(* IEC 61131-3 sources: guidance-for-physical-ai-production-designer-on-aws/source/plan2cell/examples/welding_cell_2_small/plc/codesys/head/POU, 8 files *)

(* ---- FB_Cell.st ---- *)
(*
 * FB_Cell
 * Generated by bt2plc 0.1.0 for cell welding_cell_2_small (plan bt_1790934549_welding_cell_2_small)
 *
 * Cell control for 2 robot(s): bring-up, blind homing (HOME_FOLGE), production
 * cycle (awRobotProdFolge started on every active robot; the robots run autonomously),
 * zone / permit arbitration (FB_ZoneArbiter), supervision (op index sequence, per-op
 * watchdog, zone-wait deadline, stall, program completeness), abort (stop all, drop grants,
 * rewind tickets), recovery confirmation and reset (Reset held >= 500 ms).
 *
 *   INIT -> BRINGUP -> HOMING_SELECT <-> HOMING_RUN -> READY -> START_JOBS -> RUNNING
 *        -> CYCLE_DONE -> READY ...
 *   any fault -> ABORTING -> ERROR -(bReset)-> RESETTING -> BRINGUP -> HOMING_SELECT ...
 *   abort with a robot inside its program (op index > 0, grant held, program left
 *   incomplete or away from home), or the first bring-up after INIT (head restart /
 *   download) with an active robot away from home:
 *        ... BRINGUP -> RECOVERY -(bRecoveryConfirm)-> RESETTING -> BRINGUP -> HOMING_SELECT
 *        (operator moves the robots clear in T1 first; homing is then always sequential)
 *   Start-up homing stays automatic when every active robot is at home.
 *
 * Operator: a bStop edge is latched in every state until it is consumed - abort (normal
 * states), cancel of the reset -> ERROR (INIT / RESETTING, driver Reset low), or cleared
 * (ERROR). A bReset edge in ABORTING is applied when ERROR is reached.
 *
 * Scan order: robot drivers (commands of the previous scan) -> op index tracking ->
 * faults known so far -> arbiter (this scan's inputs, no new grants after a fault) ->
 * watchdogs -> faults -> state machine -> GRANT bytes (0 when a fault is latched).
 * Op supervision runs whenever a robot's production job is commanded / running, in any
 * cell state: op index sequence, zone ops left without grant, op index 0 while running.
 *
 * Portable: one FB_VassRobot instance per robot (no FB instance arrays), timers are
 * TIME stamps of one free-running clock (_tNow).
 *)

FUNCTION_BLOCK FB_Cell
VAR_INPUT
    bEnable             : BOOL := TRUE;
    bAutoRun            : BOOL := TRUE;     (* Level: start a cycle whenever READY *)
    bStart              : BOOL;             (* Rising edge: start one cycle *)
    bStop               : BOOL;             (* Rising edge: abort (ERR_OPERATOR_STOP) *)
    bReset              : BOOL;             (* Rising edge in CS_ERROR: reset robots and cell *)
    bRecoveryConfirm    : BOOL;             (* Rising edge (from CS_ERROR on, while bRecoveryRequired): robots cleared *)
    astIn               : ARRAY[1..2] OF ST_RobotIn;    (* Robot inputs (copied from GVL_IO) *)
END_VAR

VAR_OUTPUT
    astOut              : ARRAY[1..2] OF ST_RobotOut;   (* Robot outputs (copied to GVL_IO) *)
    eState              : E_CellState;
    eError              : E_CellError;      (* First fault, ERR_NONE when OK *)
    nErrorRobot         : INT;              (* Robot of the fault, 0 = cell *)
    nErrorOp            : INT;              (* Op index of the fault, 0 = none *)
    nErrorZone          : INT;              (* Zone of the fault, 0 = none *)
    bCycleActive        : BOOL;             (* START_JOBS or RUNNING *)
    bError              : BOOL;             (* Fault latched until the reset is done *)
    bHomingRequired     : BOOL;         (* Profile vw-ks24: a robot is not at home and must be
                                           jogged there by the operator (no blind HOME Folge) *)
    bRecoveryRequired   : BOOL;             (* bRecoveryConfirm needed before homing (abort mid-cycle / start-up away from home) *)
    udiCycles           : UDINT;            (* Completed production cycles *)
    tLastCycle          : TIME;             (* Duration of the last cycle (RUNNING) *)
    aeRobotState        : ARRAY[1..2] OF E_RobotState;
    aeRobotError        : ARRAY[1..2] OF E_CellError;
    awStep              : ARRAY[1..2] OF WORD;          (* Reported op index *)
    adwReq              : ARRAY[1..2] OF DWORD;         (* REQUEST per robot *)
    adwGrant            : ARRAY[1..2] OF DWORD;         (* GRANT per robot (as sent) *)
    anDone              : ARRAY[1..2] OF INT;           (* Ops completed in this cycle *)
    anHolder            : ARRAY[1..2] OF INT;        (* Zone holder, 0 = free *)
    anTicket            : ARRAY[1..2] OF INT;        (* Next ticket per zone *)
END_VAR

VAR
    (* ========================================================================
       ROBOT DRIVERS (one instance per robot) AND ARBITER
       ======================================================================== *)
    fbRobot_R1          : FB_VassRobot;     (* 1: robot1 - kuka_robi1 (192.168.100.11) *)
    fbRobot_R2          : FB_VassRobot;     (* 2: robot2 - kuka_robi2 (192.168.100.12) *)
    fbArbiter           : FB_ZoneArbiter;

    (* ========================================================================
       CELL STATE
       ======================================================================== *)
    _eState             : E_CellState := E_CellState.CS_INIT;
    _eLastState         : E_CellState := E_CellState.CS_INIT;
    _bFault             : BOOL;             (* Fault latched (eError valid) *)
    _bPowerOn           : BOOL;             (* Robots: bring up *)
    _bArbReset          : BOOL := TRUE;     (* Arbiter reset in the next scan *)
    _bNeedRecovery      : BOOL;             (* Latched at an abort with a robot inside its program *)
    _bRecoveryHoming    : BOOL;             (* Homing after recovery: always sequential *)
    _bEngaged           : BOOL;             (* A robot is inside its production program / holds a grant *)
    _bConfirmLatch      : BOOL;             (* bRecoveryConfirm edge seen since CS_ERROR *)
    _bFirstBringup      : BOOL := TRUE;     (* First bring-up after CS_INIT: check the home poses *)
    _bStopReq           : BOOL;             (* bStop edge, latched until consumed *)
    _bResetReq          : BOOL;             (* bReset edge seen in CS_ABORTING, applied in CS_ERROR *)
    _bFaultScan         : BOOL;             (* Fault source known before the arbiter call (this scan) *)

    (* ========================================================================
       ROBOT STATUS (copied from the driver instances every scan)
       ======================================================================== *)
    _abIdle             : ARRAY[1..2] OF BOOL;
    _abBusy             : ARRAY[1..2] OF BOOL;
    _abDrvError         : ARRAY[1..2] OF BOOL;          (* Driver in RS_ERROR / RS_RESET *)
    _abJobActive        : ARRAY[1..2] OF BOOL;
    _abJobDone          : ARRAY[1..2] OF BOOL;
    _abAtHome           : ARRAY[1..2] OF BOOL;
    _abRobotError       : ARRAY[1..2] OF BOOL;          (* Robot reports Error *)
    _abProgRunning      : ARRAY[1..2] OF BOOL;          (* Robot reports ProgRunning *)
    _awLastStep         : ARRAY[1..2] OF WORD;

    (* ========================================================================
       COMMANDS TO THE ROBOT DRIVERS (used in the next scan)
       ======================================================================== *)
    _abJobCmd           : ARRAY[1..2] OF BOOL;
    _awJob              : ARRAY[1..2] OF WORD;
    _abProdCmd          : ARRAY[1..2] OF BOOL;          (* Commanded job is the production Folge *)
    _abStopCmd          : ARRAY[1..2] OF BOOL;
    _abResetCmd         : ARRAY[1..2] OF BOOL;
    _abHoming           : ARRAY[1..2] OF BOOL;

    (* ========================================================================
       PRODUCTION CYCLE SUPERVISION
       ======================================================================== *)
    _abHasJob           : ARRAY[1..2] OF BOOL;          (* Active robot with ops *)
    _abRobotOk          : ARRAY[1..2] OF BOOL;          (* Arbiter input *)
    _anDone             : ARRAY[1..2] OF INT;           (* Arbiter input: ops completed *)
    _anStepSeen         : ARRAY[1..2] OF INT;           (* Op index seen last scan (incl. 0) *)
    _anLastStep         : ARRAY[1..2] OF INT;           (* Last validated non-zero op index *)
    _abGranted          : ARRAY[1..2] OF BOOL;          (* Current zone op has been granted *)
    _abOpRun            : ARRAY[1..2] OF BOOL;          (* Op watchdog running *)
    _atOpStart          : ARRAY[1..2] OF TIME;
    _abStallRun         : ARRAY[1..2] OF BOOL;          (* Stall watchdog running *)
    _atStallStart       : ARRAY[1..2] OF TIME;
    _abZeroRun          : ARRAY[1..2] OF BOOL;          (* Op index 0 watchdog running *)
    _atZeroStart        : ARRAY[1..2] OF TIME;
    _tCycleStart        : TIME;

    (* ========================================================================
       TIME BASE / TIMERS / EDGES
       ======================================================================== *)
    _tonClock           : TON;              (* Free-running clock, restarted every hour *)
    _tClockBase         : TIME;
    _tNow               : TIME;             (* Monotonic time of this scan *)
    _tonState           : TON;              (* State timeout, restarts on every state change *)
    _tLimit             : TIME;
    _rtrigStart         : R_TRIG;
    _rtrigStop          : R_TRIG;
    _rtrigReset         : R_TRIG;
    _rtrigConfirm       : R_TRIG;

    (* ========================================================================
       SCRATCH
       ======================================================================== *)
    _eNew               : E_CellError;
    _nNewRobot          : INT;
    _nNewOp             : INT;
    _nHomeCount         : INT;
    _nDone              : INT;
    _r                  : INT;
    _iOp                : INT;
    _nStep              : INT;
    _nPrev              : INT;              (* Op index that is left *)
    _tZeroLimit         : TIME;
    _dwGrant            : DWORD;
    _bBypass            : BOOL;
    _bAll               : BOOL;
    _bSequential        : BOOL;

    (* Profile vw-ks24: interlock grant / partner release encoding *)
    _z                  : INT;
    _q                  : INT;
    _nIl                : INT;
    _nIlQ               : INT;
    _nIdx               : INT;
    _nB                 : INT;
    _nBit               : INT;
    _wBits              : WORD;
    _bGrantBit          : BOOL;
    _bPartner           : BOOL;
END_VAR

(* ---- FB_VassRobot.st ---- *)
(*
 * FB_VassRobot
 * Generated by bt2plc 0.1.0 for cell welding_cell_2_small (plan bt_1790934549_welding_cell_2_small)
 *
 * VW VASS protocol driver for ONE robot (KUKA VKRC nexxt V8.2 DIM 2 via PROFINET).
 * Portable: no pointers, no REFERENCE, no OOP - the robot IO is passed as struct
 * copies (stIn / stOut) by the caller (FB_Cell, PLC_PRG copies GVL_IO).
 *
 *   Bring-up : SAFETY_ENABLE (T_BRINGUP_LIMIT: PROFINET / PROFIsafe connection set-up)
 *              -> DRIVES_ON -> MODE_EXT -> IDLE   (T_HANDSHAKE each)
 *   Job      : WAIT_READY -> SEND (echo checked) -> START (T_START_PULSE) -> WAIT_RUNNING
 *              -> RUNNING -> DONE   (WAIT_RUNNING -> DONE if the job finished between scans)
 *              (RUNNING -> ERROR ERR_ROBOT_STOPPED only after ProgRunning and ProgFinished
 *              stayed low for T_STOP_DEBOUNCE: a robot may publish the two bits in different
 *              bus frames at the Folge end)
 *              (T_HANDSHAKE per handshake state)
 *   Abort    : STOPPING (Stop + Cancel held >= T_STOP_PULSE and until ProgRunning drops)
 *   Recovery : ERROR -> RESET (Reset held T_RESET_PULSE >= 500 ms while bCmdReset stays TRUE;
 *              bCmdReset dropped = reset cancelled -> ERROR) -> SAFETY_ENABLE
 *              (still ProgRunning after the pulse -> ERROR, ERR_STOP_TIMEOUT)
 *   Command handshake: bCmdJob is a level request (rising edge latched),
 *              bJobDone the acknowledge (cleared while bCmdJob = FALSE).
 *
 * Stop is never dropped while the robot still reports ProgRunning (also in ERROR / RESET).
 * ProgRunning outside a job (OFF, bring-up, IDLE) -> ERROR (ERR_UNEXPECTED_RUN, Stop + Cancel).
 * The zone GRANT bytes (GVL_Cell.GRANT_BYTE .. +3) are written 0 here: FB_Cell encodes
 * them after FB_ZoneArbiter has run, so a grant reaches the robot in the scan it is computed.
 *
 * Profile vw-ks24 (GVL_Cell.PROFILE_VW): the VW tech package on the robot does the Folge
 * handshake, so the signal map and the job states differ (same state names):
 *   status  : ready A9, safety A10 + A13, auto A12, home A15 (PF0), Folge end A14,
 *             echo PRG_NR_REFL A1-8, op index P_PktNr_SPS, error code VW_FEH_BIN_A
 *   commands: drives E10, Folge number PRG_NR E1-8, start SRB E9 (level), reset E26
 *   job     : SEND writes PRG_NR and waits for the echo; START holds SRB until the robot
 *             leaves home (its cycle-start point clears PF0); RUNNING waits for Folge end;
 *             DONE clears PRG_NR and waits for the Folge end to fall
 *   zones   : REQUEST bit z is synthesised as "requesting or occupying",
 *             A(80+n) OR NOT A(40+n), which is exactly the REQUEST semantics of the arbiter;
 *             the release is A(40+n) going TRUE again. There is no 4-phase handshake.
 *   stop    : no Stop/Cancel bits exist; the head drops the drives, withdraws the partner
 *             releases (the robot's online driving condition stops it on the path) and clears
 *             PRG_NR. Recovery needs manual homing (PF0), there is no blind HOME Folge.
 *)

FUNCTION_BLOCK FB_VassRobot
VAR_INPUT
    bEnable             : BOOL := TRUE;
    nRobot              : INT := 1;         (* 1-based robot index (profile vw-ks24: interlock map) *)
    bPowerOn            : BOOL;             (* Level: bring the robot up *)
    bCmdJob             : BOOL;             (* Level request (rising edge latched): run job wJobNr *)
    wJobNr              : WORD;             (* Folge number, latched at job accept *)
    bProdJob            : BOOL;             (* wJobNr is the production Folge: send PLAN_ID, track wLastStep *)
    bCmdStop            : BOOL;             (* Level: abort the active job *)
    bCmdReset           : BOOL;             (* Rising edge in RS_ERROR: reset the robot; hold until bError drops *)
    stIn                : ST_RobotIn;       (* Copy of this robot's GVL_IO inputs *)
END_VAR

VAR_OUTPUT
    stOut               : ST_RobotOut;      (* Copy to this robot's GVL_IO outputs (GRANT bytes = 0) *)
    eState              : E_RobotState;
    eError              : E_CellError;
    bIdle               : BOOL;
    bBusy               : BOOL;             (* Job, stopping or resetting *)
    bJobActive          : BOOL;             (* Job started and ProgRunning *)
    bJobDone            : BOOL;             (* Job finished (cleared while bCmdJob = FALSE) *)
    bError              : BOOL;             (* RS_ERROR or RS_RESET *)

    (* Decoded robot status *)
    bDrivesOn           : BOOL;
    bProgRunning        : BOOL;
    bAtHome             : BOOL;
    bModeExt            : BOOL;
    bRobotReady         : BOOL;
    bRobotError         : BOOL;
    bProgFinished       : BOOL;
    bJobAck             : BOOL;
    bSafetyOK           : BOOL;
    wActiveJob          : WORD;             (* Echoed job number *)
    wStep               : WORD;             (* Reported op index, 0 = no program *)
    wLastStep           : WORD;             (* Max op index of the running production job (cleared at job accept) *)
    dwZoneReq           : DWORD;            (* REQUEST DWORD: zone bits 0..30, permit bit 31 *)
    wRobotErrorCode     : WORD;
END_VAR

VAR
    _eState             : E_RobotState := E_RobotState.RS_OFF;
    _eLastState         : E_RobotState := E_RobotState.RS_OFF;
    _wJob               : WORD;             (* Job number latched at accept *)
    _bProdJob           : BOOL;             (* Latched bProdJob *)
    _bJobPending        : BOOL;             (* Job edge seen, not yet accepted *)
    _bInJob             : BOOL;
    _bUp                : BOOL;
    _bNoJob             : BOOL;             (* Off / bring-up / idle: ProgRunning is not expected *)

    (* Commands to the robot *)
    _bSafeEnable        : BOOL;
    _bDrivesOnCmd       : BOOL;
    _bExtCmd            : BOOL;
    _bStartCmd          : BOOL;
    _bStopCmd           : BOOL;
    _bCancelCmd         : BOOL;
    _bResetCmd          : BOOL;
    _bJobReqCmd         : BOOL;

    (* Timers *)
    _tonStep            : TON;              (* State timeout, restarts on every state change *)
    _tonPulse           : TON;              (* Start / stop / reset pulse width *)
    _tonStopDebounce    : TON;              (* RS_JOB_RUNNING: ProgRunning + ProgFinished low (T_STOP_DEBOUNCE) *)
    _tStepLimit         : TIME;

    (* Edge detection *)
    _rtrigJob           : R_TRIG;
    _rtrigReset         : R_TRIG;

    (* Profile vw-ks24 *)
    _bFolgeEnd          : BOOL;             (* A14 Folge end *)
    _bVwStarted         : BOOL;             (* SRB acknowledged: the robot left its home point *)
    _nIdx               : INT;              (* signal index 1..256 *)
    _nB                 : INT;              (* telegram byte of _nIdx *)
    _nBit               : INT;              (* bit of _nIdx *)
    _wTmp               : WORD;
    _bTmp               : BOOL;
    _z                  : INT;
    _n                  : INT;

    _i                  : INT;
END_VAR

(* ---- FB_ZoneArbiter.st ---- *)
(*
 * FB_ZoneArbiter
 * Generated by bt2plc 0.1.0 for cell welding_cell_2_small (plan bt_1790934549_welding_cell_2_small)
 *
 * Zone (mutex) and permit arbiter, data-driven by GVL_Cell (aTickets, anZoneFirst/Count,
 * aOps[].dwZoneMask / nPredFirst / nPredCount, aPreds).
 *
 * REQUEST / GRANT DWORD: bits 0..30 = zones 1..31, bit 31 = PERMIT (GVL_Cell.PERMIT_MASK).
 *   GP_PLANNED : a zone is granted only to its next ticket holder, only if the request
 *                equals the op's full mask and the reported op index matches the ticket.
 *   GP_FCFS    : free zones to any requester whose request equals the op mask, oldest
 *                request first, ties by robot index; zones of an older requester that
 *                waits only for occupied zones are reserved against younger ones.
 *                BT ordering is NOT preserved by the zones.
 *   PERMIT     : granted for op (r, k) iff every pred (q, j) of the op has anDone[q] >= j.
 *                Not a mutex: never held against other robots, released when bit 31 drops.
 * Both policies grant all bits of an op in the same scan (all-or-nothing).
 *
 * Checks: 4-phase handshake (op index must not change while a grant is held), release
 * only by a robot that runs OK, holder raising extra bits; request mask and ticket checks
 * are evaluated once (op index, REQUEST) has been stable for tDebounce.
 * Fail closed: any violation latches bFault and drops all grants until bReset.
 *
 * Timing uses tNow (monotonic TIME from the caller's clock), no timer instances.
 *)

FUNCTION_BLOCK FB_ZoneArbiter
VAR_INPUT
    bReset              : BOOL;             (* Level: rewind tickets, clear holders, grants and fault *)
    bEnable             : BOOL;             (* New grants allowed *)
    ePolicy             : E_GrantPolicy := E_GrantPolicy.GP_PLANNED;
    tDebounce           : TIME := T#200MS;  (* (op index, REQUEST) stable time before mask / ticket checks *)
    tNow                : TIME;             (* Monotonic time of this scan *)
    abRobotOk           : ARRAY[1..2] OF BOOL;      (* Production job running, no robot error *)
    awStep              : ARRAY[1..2] OF WORD;      (* Reported op index, 0 = none *)
    adwReq              : ARRAY[1..2] OF DWORD;     (* REQUEST DWORD *)
    anDone              : ARRAY[1..2] OF INT;       (* Ops completed per robot in this cycle *)
END_VAR

VAR_OUTPUT
    adwGrant            : ARRAY[1..2] OF DWORD;     (* GRANT DWORD per robot *)
    anHolder            : ARRAY[1..2] OF INT;    (* Robot holding the zone, 0 = free *)
    anTicket            : ARRAY[1..2] OF INT;    (* Next ticket index in GVL_Cell.aTickets *)
    bAllConsumed        : BOOL;             (* No zone held and (planned) every ticket consumed *)
    bFault              : BOOL;
    eFault              : E_CellError;
    nFaultRobot         : INT;
    nFaultZone          : INT;
END_VAR

VAR
    _udiScan            : UDINT;            (* Scan counter: request age for FCFS *)
    _audiWaitSince      : ARRAY[1..2] OF UDINT;     (* Scan of the first pending request, 0 = none *)
    _abPicked           : ARRAY[1..2] OF BOOL;
    _anGrantStep        : ARRAY[1..2] OF INT;       (* Op index at the time of the grant *)
    _awPrevStep         : ARRAY[1..2] OF WORD;
    _adwPrevReq         : ARRAY[1..2] OF DWORD;
    _atChange           : ARRAY[1..2] OF TIME;      (* tNow of the last (op index, REQUEST) change *)
    _abStable           : ARRAY[1..2] OF BOOL;
    _eNew               : E_CellError;
    _nNewRobot          : INT;
    _nNewZone           : INT;
    _k                  : INT;
    _r                  : INT;
    _rr                 : INT;
    _rSel               : INT;
    _z                  : INT;
    _p                  : INT;
    _q                  : INT;
    _iOp                : INT;
    _nStep              : INT;
    _nTicket            : INT;
    _nLastTicket        : INT;
    _nPredFirst         : INT;
    _nPredLast          : INT;
    _dwBit              : DWORD;
    _dwExp              : DWORD;            (* Expected REQUEST of the reported op *)
    _dwZones            : DWORD;            (* Zone bits of _dwExp (permit bit removed) *)
    _dwReserved         : DWORD;            (* FCFS: zones reserved by older requesters this scan *)
    _bOk                : BOOL;             (* All zones of the op grantable *)
    _bPermitOk          : BOOL;             (* All permit predecessors done *)
    _bPending           : BOOL;
END_VAR

(* ---- FB_Cell_Body.st ---- *)
(*
 * FB_Cell - Implementation
 *)

IF NOT bEnable THEN
    _eState := E_CellState.CS_INIT;
END_IF

(* ============================================================================
   TIME BASE / EDGES
   ============================================================================ *)
_tonClock(IN := TRUE, PT := T#1H);
_tNow := _tClockBase + _tonClock.ET;
IF _tonClock.Q THEN
    _tClockBase := _tNow;
    _tonClock(IN := FALSE);
    _tonClock(IN := TRUE, PT := T#1H);
END_IF

_rtrigStart(CLK := bStart);
_rtrigStop(CLK := bStop);
_rtrigReset(CLK := bReset);
_rtrigConfirm(CLK := bRecoveryConfirm);

(* Operator stop: latched in every state until consumed (abort, cancelled reset, CS_ERROR);
   it also cancels a reset that is pending from CS_ABORTING *)
IF _rtrigStop.Q THEN
    _bStopReq := TRUE;
    _bResetReq := FALSE;
END_IF

FOR _r := 1 TO GVL_Cell.N_ROBOTS DO
    _abHasJob[_r] := GVL_Cell.abRobotActive[_r] AND (GVL_Cell.anRobotOpCount[_r] > 0);
END_FOR

(* ============================================================================
   ROBOT DRIVERS (commands from the previous scan; GRANT bytes are added below)
   ============================================================================ *)

(* 1: R1 - robot1 *)
fbRobot_R1(
    bEnable     := bEnable,
    bPowerOn    := _bPowerOn,
    bCmdJob     := _abJobCmd[1],
    wJobNr      := _awJob[1],
    bProdJob    := _abProdCmd[1],
    bCmdStop    := _abStopCmd[1],
    bCmdReset   := _abResetCmd[1],
    nRobot      := 1,
    stIn        := astIn[1]);
astOut[1]         := fbRobot_R1.stOut;
aeRobotState[1]   := fbRobot_R1.eState;
aeRobotError[1]   := fbRobot_R1.eError;
awStep[1]         := fbRobot_R1.wStep;
adwReq[1]         := fbRobot_R1.dwZoneReq;
_awLastStep[1]    := fbRobot_R1.wLastStep;
_abIdle[1]        := fbRobot_R1.bIdle;
_abBusy[1]        := fbRobot_R1.bBusy;
_abDrvError[1]    := fbRobot_R1.bError;
_abJobActive[1]   := fbRobot_R1.bJobActive;
_abJobDone[1]     := fbRobot_R1.bJobDone;
_abAtHome[1]      := fbRobot_R1.bAtHome;
_abRobotError[1]  := fbRobot_R1.bRobotError;
_abProgRunning[1] := fbRobot_R1.bProgRunning;

(* 2: R2 - robot2 *)
fbRobot_R2(
    bEnable     := bEnable,
    bPowerOn    := _bPowerOn,
    bCmdJob     := _abJobCmd[2],
    wJobNr      := _awJob[2],
    bProdJob    := _abProdCmd[2],
    bCmdStop    := _abStopCmd[2],
    bCmdReset   := _abResetCmd[2],
    nRobot      := 2,
    stIn        := astIn[2]);
astOut[2]         := fbRobot_R2.stOut;
aeRobotState[2]   := fbRobot_R2.eState;
aeRobotError[2]   := fbRobot_R2.eError;
awStep[2]         := fbRobot_R2.wStep;
adwReq[2]         := fbRobot_R2.dwZoneReq;
_awLastStep[2]    := fbRobot_R2.wLastStep;
_abIdle[2]        := fbRobot_R2.bIdle;
_abBusy[2]        := fbRobot_R2.bBusy;
_abDrvError[2]    := fbRobot_R2.bError;
_abJobActive[2]   := fbRobot_R2.bJobActive;
_abJobDone[2]     := fbRobot_R2.bJobDone;
_abAtHome[2]      := fbRobot_R2.bAtHome;
_abRobotError[2]  := fbRobot_R2.bRobotError;
_abProgRunning[2] := fbRobot_R2.bProgRunning;

(* A robot inside its production program or holding a grant (previous scan's commands):
   inside an op, between two ops, finished with an incomplete program, or left the
   home pose during the current cycle *)
_bEngaged := FALSE;
FOR _r := 1 TO GVL_Cell.N_ROBOTS DO
    IF _abJobCmd[_r] AND _abProdCmd[_r] THEN
        IF awStep[_r] <> WORD#0 THEN
            _bEngaged := TRUE;
        ELSIF (_awLastStep[_r] <> WORD#0) AND NOT _abJobDone[_r] THEN
            _bEngaged := TRUE;
        ELSIF _abJobDone[_r] AND (WORD_TO_INT(_awLastStep[_r]) <> GVL_Cell.anRobotOpCount[_r]) THEN
            _bEngaged := TRUE;
        ELSIF NOT _abAtHome[_r]
              AND ((_awLastStep[_r] <> WORD#0) OR (_anLastStep[_r] <> 0) OR _abJobActive[_r]) THEN
            _bEngaged := TRUE;
        END_IF
    END_IF
    IF fbArbiter.adwGrant[_r] <> DWORD#0 THEN
        _bEngaged := TRUE;
    END_IF
END_FOR

(* ============================================================================
   OP INDEX TRACKING (production job commanded, any cell state)
   The index must advance by exactly +1. The op that is left (also at the job end,
   index -> 0) must have been granted if it has a zone / permit mask (both policies).
   Index 0 while the program runs is valid only before the first / after the last op.
   ============================================================================ *)
_eNew := E_CellError.ERR_NONE;
_nNewRobot := 0;
_nNewOp := 0;
FOR _r := 1 TO GVL_Cell.N_ROBOTS DO
    IF _abJobCmd[_r] AND _abProdCmd[_r] THEN
        _nStep := WORD_TO_INT(awStep[_r]);
        IF _nStep <> _anStepSeen[_r] THEN
            _nPrev := _anStepSeen[_r];
            _bBypass := FALSE;
            IF (_nPrev >= 1) AND (_nPrev <= GVL_Cell.anRobotOpCount[_r]) AND NOT _abGranted[_r] THEN
                _iOp := GVL_Cell.anRobotFirstOp[_r] + _nPrev - 1;
                IF GVL_Cell.aOps[_iOp].dwZoneMask <> DWORD#0 THEN
                    _bBypass := TRUE;               (* zone / permit op left without a grant *)
                END_IF
            END_IF
            IF _bBypass THEN
                IF _eNew = E_CellError.ERR_NONE THEN
                    _eNew := E_CellError.ERR_ZONE_BYPASSED;
                    _nNewRobot := _r;
                    _nNewOp := _nPrev;
                END_IF
            ELSIF _nStep <> 0 THEN
                IF (_nStep = _anLastStep[_r] + 1) AND (_nStep <= GVL_Cell.anRobotOpCount[_r]) THEN
                    _anLastStep[_r] := _nStep;
                ELSIF _eNew = E_CellError.ERR_NONE THEN
                    _eNew := E_CellError.ERR_STEP_SEQUENCE;
                    _nNewRobot := _r;
                    _nNewOp := _nStep;
                END_IF
            END_IF
            _anStepSeen[_r] := _nStep;
            _abGranted[_r] := FALSE;
            _abOpRun[_r] := FALSE;
            _abStallRun[_r] := FALSE;
            _abZeroRun[_r] := FALSE;
        END_IF

        (* index 0 while the program runs, between two ops *)
        IF _abJobActive[_r] AND (_nStep = 0) AND (_anLastStep[_r] > 0)
           AND (_anLastStep[_r] < GVL_Cell.anRobotOpCount[_r])
           AND (_eNew = E_CellError.ERR_NONE) THEN
            _eNew := E_CellError.ERR_STEP_SEQUENCE;
            _nNewRobot := _r;
            _nNewOp := 0;
        END_IF

        (* ops completed (permit predecessors): validated index - 1, all at job done *)
        IF _abJobDone[_r] AND (_anLastStep[_r] = GVL_Cell.anRobotOpCount[_r]) THEN
            _nDone := GVL_Cell.anRobotOpCount[_r];
        ELSIF _anLastStep[_r] > 0 THEN
            _nDone := _anLastStep[_r] - 1;
        ELSE
            _nDone := 0;
        END_IF
        _anDone[_r] := MAX(_anDone[_r], _nDone);
    END_IF
END_FOR

(* ============================================================================
   ZONE ARBITER (this scan's robot inputs)
   No new grants in a scan in which the cell already knows it will abort:
   driver error, latched operator stop, latched fault, supervision fault above.
   ============================================================================ *)
_bFaultScan := _bFault OR _bStopReq OR (_eNew <> E_CellError.ERR_NONE);
FOR _r := 1 TO GVL_Cell.N_ROBOTS DO
    _abRobotOk[_r] := _abJobActive[_r] AND _abJobCmd[_r] AND _abProdCmd[_r] AND NOT _abRobotError[_r];
    IF _abDrvError[_r] THEN
        _bFaultScan := TRUE;
    END_IF
END_FOR
fbArbiter(
    bReset      := _bArbReset,
    bEnable     := ((_eState = E_CellState.CS_START_JOBS) OR (_eState = E_CellState.CS_RUNNING))
                   AND NOT _bFaultScan,
    ePolicy     := GVL_Cell.GRANT_POLICY,
    tDebounce   := GVL_Cell.T_MISMATCH_DEBOUNCE,
    tNow        := _tNow,
    abRobotOk   := _abRobotOk,
    awStep      := awStep,
    adwReq      := adwReq,
    anDone      := _anDone);
_bArbReset := FALSE;

(* ============================================================================
   WATCHDOGS (production job running, any cell state)
   op watchdog from the step change (mask 0) or from the grant; stall; zone wait;
   op index 0: T_HANDSHAKE before the first op, MAX(last op tLimit, T_HANDSHAKE)
   after the last op
   ============================================================================ *)
FOR _r := 1 TO GVL_Cell.N_ROBOTS DO
    IF _abJobCmd[_r] AND _abProdCmd[_r] AND _abJobActive[_r] THEN
        _nStep := _anStepSeen[_r];
        IF (_nStep >= 1) AND (_nStep <= GVL_Cell.anRobotOpCount[_r]) THEN
            _iOp := GVL_Cell.anRobotFirstOp[_r] + _nStep - 1;
            IF GVL_Cell.aOps[_iOp].dwZoneMask = DWORD#0 THEN
                IF NOT _abOpRun[_r] THEN
                    _abOpRun[_r] := TRUE;
                    _atOpStart[_r] := _tNow;
                END_IF
            ELSE
                IF fbArbiter.adwGrant[_r] <> DWORD#0 THEN
                    _abGranted[_r] := TRUE;
                END_IF
                IF _abGranted[_r] AND NOT _abOpRun[_r] THEN
                    _abOpRun[_r] := TRUE;
                    _atOpStart[_r] := _tNow;
                END_IF

                (* zone op with neither REQUEST nor grant *)
                IF NOT _abGranted[_r] AND (adwReq[_r] = DWORD#0) THEN
                    IF NOT _abStallRun[_r] THEN
                        _abStallRun[_r] := TRUE;
                        _atStallStart[_r] := _tNow;
                    ELSIF ((_tNow - _atStallStart[_r]) >= GVL_Cell.T_HANDSHAKE)
                          AND (_eNew = E_CellError.ERR_NONE) THEN
                        _eNew := E_CellError.ERR_ROBOT_STALLED;
                        _nNewRobot := _r;
                        _nNewOp := _nStep;
                    END_IF
                ELSE
                    _abStallRun[_r] := FALSE;
                END_IF

                (* zone wait past the deadline (measured since the cycle started RUNNING) *)
                IF NOT _abGranted[_r] AND (adwReq[_r] <> DWORD#0)
                   AND (_eState = E_CellState.CS_RUNNING)
                   AND ((_tNow - _tCycleStart) > GVL_Cell.aOps[_iOp].tZoneDeadline)
                   AND (_eNew = E_CellError.ERR_NONE) THEN
                    _eNew := E_CellError.ERR_ZONE_WAIT_TIMEOUT;
                    _nNewRobot := _r;
                    _nNewOp := _nStep;
                END_IF
            END_IF

            IF _abOpRun[_r] AND ((_tNow - _atOpStart[_r]) >= GVL_Cell.aOps[_iOp].tLimit)
               AND (_eNew = E_CellError.ERR_NONE) THEN
                _eNew := E_CellError.ERR_OP_WATCHDOG;
                _nNewRobot := _r;
                _nNewOp := _nStep;
            END_IF
        ELSIF _nStep = 0 THEN
            (* program running without an op: before the first / after the last op *)
            IF NOT _abZeroRun[_r] THEN
                _abZeroRun[_r] := TRUE;
                _atZeroStart[_r] := _tNow;
            END_IF
            _tZeroLimit := GVL_Cell.T_HANDSHAKE;
            IF (_anLastStep[_r] >= 1) AND (_anLastStep[_r] = GVL_Cell.anRobotOpCount[_r]) THEN
                _iOp := GVL_Cell.anRobotFirstOp[_r] + _anLastStep[_r] - 1;
                IF GVL_Cell.aOps[_iOp].tLimit > _tZeroLimit THEN
                    _tZeroLimit := GVL_Cell.aOps[_iOp].tLimit;
                END_IF
            END_IF
            IF ((_tNow - _atZeroStart[_r]) >= _tZeroLimit) AND (_eNew = E_CellError.ERR_NONE) THEN
                _eNew := E_CellError.ERR_ROBOT_STALLED;
                _nNewRobot := _r;
                _nNewOp := 0;
            END_IF
        END_IF
    ELSE
        _abZeroRun[_r] := FALSE;
    END_IF
END_FOR

(* ============================================================================
   FAULT COLLECTION (first wins: robot > supervision > arbiter > operator)
   ============================================================================ *)
IF (_eState <> E_CellState.CS_INIT) AND (_eState <> E_CellState.CS_ABORTING)
   AND (_eState <> E_CellState.CS_ERROR) AND (_eState <> E_CellState.CS_RESETTING) THEN
    FOR _r := 1 TO GVL_Cell.N_ROBOTS DO
        IF _abDrvError[_r] AND NOT _bFault AND (_eState <> E_CellState.CS_RECOVERY) THEN
            _bFault := TRUE;
            eError := aeRobotError[_r];
            nErrorRobot := _r;
            nErrorOp := WORD_TO_INT(awStep[_r]);
            nErrorZone := 0;
        END_IF
    END_FOR
    IF (_eNew <> E_CellError.ERR_NONE) AND NOT _bFault THEN
        _bFault := TRUE;
        eError := _eNew;
        nErrorRobot := _nNewRobot;
        nErrorOp := _nNewOp;
        nErrorZone := 0;
    END_IF
    IF fbArbiter.bFault AND NOT _bFault THEN
        _bFault := TRUE;
        eError := fbArbiter.eFault;
        nErrorRobot := fbArbiter.nFaultRobot;
        nErrorOp := 0;
        IF (fbArbiter.nFaultRobot >= 1) AND (fbArbiter.nFaultRobot <= GVL_Cell.N_ROBOTS) THEN
            nErrorOp := WORD_TO_INT(awStep[fbArbiter.nFaultRobot]);
        END_IF
        nErrorZone := fbArbiter.nFaultZone;
    END_IF
    IF _bStopReq THEN
        _bStopReq := FALSE;                 (* consumed by this abort *)
        IF NOT _bFault THEN
            _bFault := TRUE;
            eError := E_CellError.ERR_OPERATOR_STOP;
            nErrorRobot := 0;
            nErrorOp := 0;
            nErrorZone := 0;
        END_IF
    END_IF
    IF _bFault THEN
        _eState := E_CellState.CS_ABORTING;
    END_IF
END_IF

(* ============================================================================
   STATE TIMER (after the transitions above: a new state starts with a fresh timer)
   ============================================================================ *)
IF _eState <> _eLastState THEN
    IF _eState = E_CellState.CS_ABORTING THEN
        _bConfirmLatch := FALSE;
        IF _bEngaged THEN
            _bNeedRecovery := TRUE;         (* aborted with a robot inside its program *)
        END_IF
    END_IF
    _tonState(IN := FALSE);
    _eLastState := _eState;
END_IF
CASE _eState OF
E_CellState.CS_HOMING_RUN:
    _tLimit := GVL_Cell.T_HOME_LIMIT;
E_CellState.CS_START_JOBS:
    _tLimit := GVL_Cell.T_START_LIMIT;
E_CellState.CS_CYCLE_DONE:
    _tLimit := GVL_Cell.T_CYCLE_PAUSE;
E_CellState.CS_ABORTING, E_CellState.CS_RESETTING:
    _tLimit := GVL_Cell.T_ABORT_LIMIT;
ELSE
    _tLimit := T#24H;
END_CASE
_tonState(IN := TRUE, PT := _tLimit);

(* Recovery confirm: accepted once the robots are stopped (CS_ERROR on), used in CS_RECOVERY *)
IF _rtrigConfirm.Q AND _bNeedRecovery
   AND ((_eState = E_CellState.CS_ERROR) OR (_eState = E_CellState.CS_RESETTING)
        OR (_eState = E_CellState.CS_BRINGUP) OR (_eState = E_CellState.CS_RECOVERY)) THEN
    _bConfirmLatch := TRUE;
END_IF

(* ============================================================================
   STATE MACHINE
   ============================================================================ *)
CASE _eState OF

E_CellState.CS_INIT:
    _bPowerOn := FALSE;
    _bArbReset := TRUE;
    _bFirstBringup := TRUE;                 (* head start / restart: robot poses unknown *)
    FOR _r := 1 TO GVL_Cell.N_ROBOTS DO
        _abJobCmd[_r] := FALSE;
        _abProdCmd[_r] := FALSE;
        _abStopCmd[_r] := FALSE;
        _abResetCmd[_r] := FALSE;
        _abHoming[_r] := FALSE;
    END_FOR
    IF bEnable THEN
        IF _bStopReq THEN
            (* operator stop before the start-up: no automatic bring-up *)
            _bStopReq := FALSE;
            _bResetReq := FALSE;
            _bFault := TRUE;
            eError := E_CellError.ERR_OPERATOR_STOP;
            nErrorRobot := 0;
            nErrorOp := 0;
            nErrorZone := 0;
            _eState := E_CellState.CS_ERROR;
        ELSE
            _eState := E_CellState.CS_BRINGUP;
        END_IF
    END_IF

E_CellState.CS_BRINGUP:
    _bPowerOn := TRUE;
    _bAll := TRUE;
    FOR _r := 1 TO GVL_Cell.N_ROBOTS DO
        IF NOT _abIdle[_r] THEN
            _bAll := FALSE;
        END_IF
    END_FOR
    IF _bAll THEN
        IF _bFirstBringup THEN
            (* first bring-up after INIT: any robot away from home (also an idle one)
               may stand anywhere in the shared space (head restart / download mid-cycle) *)
            _bFirstBringup := FALSE;
            FOR _r := 1 TO GVL_Cell.N_ROBOTS DO
                IF NOT _abAtHome[_r] AND NOT _bNeedRecovery THEN
                    _bNeedRecovery := TRUE;
                    _bConfirmLatch := FALSE;
                END_IF
            END_FOR
        END_IF
        IF _bNeedRecovery THEN
            _eState := E_CellState.CS_RECOVERY;
        ELSE
            _eState := E_CellState.CS_HOMING_SELECT;
        END_IF
    END_IF

E_CellState.CS_RECOVERY:
    (* robots may be anywhere inside the shared space: the operator moves them
       clear (T1, driver errors are ignored here) and confirms; then the drivers
       are reset, brought up again and blind homing runs one robot at a time *)
    IF _bConfirmLatch THEN
        _bConfirmLatch := FALSE;
        _bNeedRecovery := FALSE;
        _bRecoveryHoming := TRUE;
        _eState := E_CellState.CS_RESETTING;
    END_IF

E_CellState.CS_HOMING_SELECT:
    IF GVL_Cell.PROFILE_VW THEN
        (* VW cell.src starts a Folge only once the robot reports PF0, and there is no blind
           home Folge: wait for the operator to jog every robot home (ERR_HOME_FAILED on
           T_HOME_LIMIT tells which robot is not at home). *)
        _bAll := TRUE;
        FOR _r := 1 TO GVL_Cell.N_ROBOTS DO
            IF NOT _abAtHome[_r] THEN
                _bAll := FALSE;
                bHomingRequired := TRUE;
            END_IF
        END_FOR
        IF _bAll THEN
            bHomingRequired := FALSE;
            _bRecoveryHoming := FALSE;
            _eState := E_CellState.CS_READY;
        ELSIF _tonState.Q THEN
            _bFault := TRUE;
            eError := E_CellError.ERR_HOME_FAILED;
            nErrorRobot := 0;
            FOR _r := GVL_Cell.N_ROBOTS TO 1 BY -1 DO
                IF NOT _abAtHome[_r] THEN
                    nErrorRobot := _r;
                END_IF
            END_FOR
            nErrorOp := 0;
            nErrorZone := 0;
            _eState := E_CellState.CS_ERROR;
        END_IF
    ELSE
        _bSequential := GVL_Cell.HOME_SEQUENTIAL OR _bRecoveryHoming;
        _nHomeCount := 0;
        FOR _r := 1 TO GVL_Cell.N_ROBOTS DO
            _abHoming[_r] := FALSE;
            IF NOT _abAtHome[_r] AND (NOT _bSequential OR (_nHomeCount = 0)) THEN
                _abHoming[_r] := TRUE;
                _awJob[_r] := GVL_Cell.HOME_FOLGE;
                _abProdCmd[_r] := FALSE;
                _nHomeCount := _nHomeCount + 1;
            END_IF
        END_FOR
        IF _nHomeCount = 0 THEN
            _bRecoveryHoming := FALSE;
            _eState := E_CellState.CS_READY;
        ELSE
            _eState := E_CellState.CS_HOMING_RUN;
        END_IF
    END_IF

E_CellState.CS_HOMING_RUN:
    _bAll := TRUE;
    FOR _r := 1 TO GVL_Cell.N_ROBOTS DO
        IF _abHoming[_r] THEN
            _abJobCmd[_r] := TRUE;
            IF NOT _abJobDone[_r] THEN
                _bAll := FALSE;
            ELSIF NOT _abAtHome[_r] AND NOT _bFault THEN
                _bFault := TRUE;
                eError := E_CellError.ERR_HOME_FAILED;
                nErrorRobot := _r;
                nErrorOp := 0;
                nErrorZone := 0;
            END_IF
        END_IF
    END_FOR
    IF _bFault THEN
        _eState := E_CellState.CS_ABORTING;
    ELSIF _bAll THEN
        FOR _r := 1 TO GVL_Cell.N_ROBOTS DO
            IF _abHoming[_r] THEN
                _abJobCmd[_r] := FALSE;
                _abHoming[_r] := FALSE;
            END_IF
        END_FOR
        _eState := E_CellState.CS_HOMING_SELECT;
    ELSIF _tonState.Q THEN
        _bFault := TRUE;
        eError := E_CellError.ERR_HOME_FAILED;
        nErrorRobot := 0;
        FOR _r := GVL_Cell.N_ROBOTS TO 1 BY -1 DO
            IF _abHoming[_r] AND NOT _abJobDone[_r] THEN
                nErrorRobot := _r;
            END_IF
        END_FOR
        nErrorOp := 0;
        nErrorZone := 0;
        _eState := E_CellState.CS_ABORTING;
    END_IF

E_CellState.CS_READY:
    IF _rtrigStart.Q OR bAutoRun THEN
        _bAll := TRUE;
        FOR _r := 1 TO GVL_Cell.N_ROBOTS DO
            IF _abHasJob[_r] AND NOT _abAtHome[_r] THEN
                _bAll := FALSE;             (* programs start at the home pose *)
            END_IF
        END_FOR
        IF _bAll THEN
            _bArbReset := TRUE;             (* rewind tickets for this cycle *)
            FOR _r := 1 TO GVL_Cell.N_ROBOTS DO
                _anStepSeen[_r] := 0;
                _anLastStep[_r] := 0;
                _anDone[_r] := 0;
                _abGranted[_r] := FALSE;
                _abOpRun[_r] := FALSE;
                _abStallRun[_r] := FALSE;
                _abZeroRun[_r] := FALSE;
                _abProdCmd[_r] := FALSE;
                IF _abHasJob[_r] THEN
                    _awJob[_r] := GVL_Cell.awRobotProdFolge[_r];
                    _abProdCmd[_r] := TRUE;
                END_IF
            END_FOR
            _eState := E_CellState.CS_START_JOBS;
        ELSE
            _eState := E_CellState.CS_HOMING_SELECT;
        END_IF
    END_IF

E_CellState.CS_START_JOBS:
    _bAll := TRUE;
    FOR _r := 1 TO GVL_Cell.N_ROBOTS DO
        IF _abHasJob[_r] THEN
            _abJobCmd[_r] := TRUE;
            IF NOT (_abJobActive[_r] OR _abJobDone[_r]) THEN
                _bAll := FALSE;
            END_IF
        END_IF
    END_FOR
    IF _bAll THEN
        _tCycleStart := _tNow;
        _eState := E_CellState.CS_RUNNING;
    ELSIF _tonState.Q THEN
        _bFault := TRUE;
        eError := E_CellError.ERR_START_TIMEOUT;
        nErrorRobot := 0;
        FOR _r := GVL_Cell.N_ROBOTS TO 1 BY -1 DO
            IF _abHasJob[_r] AND NOT (_abJobActive[_r] OR _abJobDone[_r]) THEN
                nErrorRobot := _r;
            END_IF
        END_FOR
        nErrorOp := 0;
        nErrorZone := 0;
        _eState := E_CellState.CS_ABORTING;
    END_IF

E_CellState.CS_RUNNING:
    _bAll := TRUE;
    FOR _r := 1 TO GVL_Cell.N_ROBOTS DO
        IF _abHasJob[_r] THEN
            IF NOT _abJobDone[_r] THEN
                _bAll := FALSE;
            ELSIF (WORD_TO_INT(_awLastStep[_r]) <> GVL_Cell.anRobotOpCount[_r]) AND NOT _bFault THEN
                _bFault := TRUE;
                eError := E_CellError.ERR_PROGRAM_INCOMPLETE;
                nErrorRobot := _r;
                nErrorOp := WORD_TO_INT(_awLastStep[_r]);
                nErrorZone := 0;
            END_IF
        END_IF
    END_FOR
    IF _bFault THEN
        _eState := E_CellState.CS_ABORTING;
    ELSIF _bAll THEN
        IF NOT fbArbiter.bAllConsumed THEN
            _bFault := TRUE;
            eError := E_CellError.ERR_TICKETS_LEFT;
            nErrorRobot := 0;
            nErrorOp := 0;
            nErrorZone := 0;
            _eState := E_CellState.CS_ABORTING;
        ELSE
            FOR _r := 1 TO GVL_Cell.N_ROBOTS DO
                _abJobCmd[_r] := FALSE;
            END_FOR
            udiCycles := udiCycles + 1;
            tLastCycle := _tNow - _tCycleStart;
            _eState := E_CellState.CS_CYCLE_DONE;
        END_IF
    END_IF

E_CellState.CS_CYCLE_DONE:
    IF _tonState.Q THEN
        _eState := E_CellState.CS_READY;
    END_IF

E_CellState.CS_ABORTING:
    _bArbReset := TRUE;                     (* drop all grants, rewind tickets *)
    _bAll := TRUE;
    FOR _r := 1 TO GVL_Cell.N_ROBOTS DO
        _abJobCmd[_r] := FALSE;
        _abHoming[_r] := FALSE;
        _abStopCmd[_r] := TRUE;
        IF _abBusy[_r] THEN
            _bAll := FALSE;
        END_IF
    END_FOR
    IF _rtrigReset.Q AND NOT _rtrigStop.Q THEN
        _bResetReq := TRUE;                 (* applied once CS_ERROR is reached *)
        _bStopReq := FALSE;                 (* the abort in progress already stops *)
    END_IF
    IF _bAll OR _tonState.Q THEN
        _eState := E_CellState.CS_ERROR;
    END_IF

E_CellState.CS_ERROR:
    _bArbReset := TRUE;
    FOR _r := 1 TO GVL_Cell.N_ROBOTS DO
        _abStopCmd[_r] := FALSE;            (* drivers keep Stop while a robot still runs *)
        _abResetCmd[_r] := FALSE;           (* re-arm the reset edges *)
    END_FOR
    IF _bStopReq THEN
        _bStopReq := FALSE;                 (* already stopped *)
        _bResetReq := FALSE;
    ELSIF _rtrigReset.Q OR _bResetReq THEN
        _bResetReq := FALSE;
        _eState := E_CellState.CS_RESETTING;
    END_IF

E_CellState.CS_RESETTING:
    IF _bStopReq THEN
        (* operator stop cancels the reset: driver Reset low, no bring-up / homing *)
        _bStopReq := FALSE;
        _bResetReq := FALSE;
        FOR _r := 1 TO GVL_Cell.N_ROBOTS DO
            _abResetCmd[_r] := FALSE;
        END_FOR
        IF _bRecoveryHoming THEN
            _bRecoveryHoming := FALSE;
            _bNeedRecovery := TRUE;         (* confirm again after the next reset *)
        END_IF
        _bConfirmLatch := FALSE;
        _bFault := TRUE;
        eError := E_CellError.ERR_OPERATOR_STOP;
        nErrorRobot := 0;
        nErrorOp := 0;
        nErrorZone := 0;
        _eState := E_CellState.CS_ERROR;
    ELSE
        _bAll := TRUE;
        FOR _r := 1 TO GVL_Cell.N_ROBOTS DO
            _abResetCmd[_r] := _abDrvError[_r];
            IF _abDrvError[_r] OR _abBusy[_r] OR _abProgRunning[_r] THEN
                _bAll := FALSE;
            END_IF
        END_FOR
        IF _bAll THEN
            FOR _r := 1 TO GVL_Cell.N_ROBOTS DO
                _abResetCmd[_r] := FALSE;
                _abProdCmd[_r] := FALSE;
            END_FOR
            _bFault := FALSE;
            eError := E_CellError.ERR_NONE;
            nErrorRobot := 0;
            nErrorOp := 0;
            nErrorZone := 0;
            _bArbReset := TRUE;
            _eState := E_CellState.CS_BRINGUP;  (* then recovery (if needed) or blind homing *)
        ELSIF _tonState.Q THEN
            IF NOT _bFault THEN                 (* reset after a recovery confirm failed *)
                _bFault := TRUE;
                eError := E_CellError.ERR_RESET_FAILED;
                nErrorRobot := 0;
                FOR _r := GVL_Cell.N_ROBOTS TO 1 BY -1 DO
                    IF _abDrvError[_r] OR _abBusy[_r] OR _abProgRunning[_r] THEN
                        nErrorRobot := _r;
                    END_IF
                END_FOR
                nErrorOp := 0;
                nErrorZone := 0;
            END_IF
            _eState := E_CellState.CS_ERROR;
        END_IF
    END_IF

END_CASE

(* ============================================================================
   GRANT BYTES (PLC -> robot, DWORD LE): non-zero only while the job runs and no
   fault is latched (also covers faults decided after the arbiter in this scan)
   ============================================================================ *)
FOR _r := 1 TO GVL_Cell.N_ROBOTS DO
    IF _abJobActive[_r] AND NOT _bFault AND NOT _bFaultScan THEN
        _dwGrant := fbArbiter.adwGrant[_r];
    ELSE
        _dwGrant := DWORD#0;
    END_IF
    adwGrant[_r] := _dwGrant;
    IF GVL_Cell.PROFILE_VW THEN
        (* Per interlock n of robot r: grant E(80+n) = the arbiter's zone bit, partner release
           E(40+n) = AND of the releases A(40+n) of the other members of that zone (the robot
           waits for it before it enters, and its online driving condition keeps watching it). *)
        FOR _z := 1 TO GVL_Cell.N_ZONES DO
            _nIl := GVL_Cell.anInterlock[(_r - 1) * GVL_Cell.N_ZONES + _z];
            IF (_nIl >= 1) AND (_nIl <= 16) THEN
                _bGrantBit := (_dwGrant AND SHL(DWORD#1, _z - 1)) <> DWORD#0;
                _bPartner := TRUE;
                FOR _q := 1 TO GVL_Cell.N_ROBOTS DO
                    IF _q <> _r THEN
                        _nIlQ := GVL_Cell.anInterlock[(_q - 1) * GVL_Cell.N_ZONES + _z];
                        IF (_nIlQ >= 1) AND (_nIlQ <= 16) THEN
                            _nIdx := GVL_Cell.VW_REL_OUT + _nIlQ - 1;
                            _nB := (_nIdx - 1) / 8;
                            _nBit := (_nIdx - 1) MOD 8;
                            IF (SHR(BYTE_TO_WORD(astIn[_q].aVassIn[_nB]), _nBit) AND WORD#1) = WORD#0 THEN
                                _bPartner := FALSE;
                            END_IF
                        END_IF
                    END_IF
                END_FOR
                _nIdx := GVL_Cell.VW_REQ_OUT + _nIl - 1;
                _nB := (_nIdx - 1) / 8;
                _nBit := (_nIdx - 1) MOD 8;
                IF _bGrantBit THEN
                    _wBits := BYTE_TO_WORD(astOut[_r].aVassOut[_nB]) OR SHL(WORD#1, _nBit);
                    astOut[_r].aVassOut[_nB] := WORD_TO_BYTE(_wBits);
                END_IF
                _nIdx := GVL_Cell.VW_REL_OUT + _nIl - 1;
                _nB := (_nIdx - 1) / 8;
                _nBit := (_nIdx - 1) MOD 8;
                IF _bPartner AND NOT _bFault AND NOT _bFaultScan THEN
                    _wBits := BYTE_TO_WORD(astOut[_r].aVassOut[_nB]) OR SHL(WORD#1, _nBit);
                    astOut[_r].aVassOut[_nB] := WORD_TO_BYTE(_wBits);
                END_IF
            END_IF
        END_FOR
    ELSE
        astOut[_r].aVassOut[GVL_Cell.GRANT_BYTE]     := DWORD_TO_BYTE(_dwGrant AND DWORD#16#FF);
        astOut[_r].aVassOut[GVL_Cell.GRANT_BYTE + 1] := DWORD_TO_BYTE(SHR(_dwGrant, 8) AND DWORD#16#FF);
        astOut[_r].aVassOut[GVL_Cell.GRANT_BYTE + 2] := DWORD_TO_BYTE(SHR(_dwGrant, 16) AND DWORD#16#FF);
        astOut[_r].aVassOut[GVL_Cell.GRANT_BYTE + 3] := DWORD_TO_BYTE(SHR(_dwGrant, 24) AND DWORD#16#FF);
    END_IF
END_FOR

(* ============================================================================
   OUTPUTS
   ============================================================================ *)
eState := _eState;
bError := _bFault;
bCycleActive := (_eState = E_CellState.CS_START_JOBS) OR (_eState = E_CellState.CS_RUNNING);
bRecoveryRequired := _bNeedRecovery;
anHolder := fbArbiter.anHolder;
anTicket := fbArbiter.anTicket;
anDone := _anDone;

(* ---- FB_VassRobot_Body.st ---- *)
(*
 * FB_VassRobot - Implementation
 * Reads the robot status from stIn, writes the commands to stOut.
 *)

IF NOT bEnable THEN
    FOR _i := 0 TO 31 DO
        stOut.aVassOut[_i] := BYTE#0;
    END_FOR
    FOR _i := 0 TO 7 DO
        stOut.abySafeOut[_i] := BYTE#0;
    END_FOR
    _eState := E_RobotState.RS_OFF;
    _eLastState := E_RobotState.RS_OFF;
    _bJobPending := FALSE;
    eState := _eState;
    eError := E_CellError.ERR_NONE;
    bIdle := FALSE;
    bBusy := FALSE;
    bJobActive := FALSE;
    bJobDone := FALSE;
    bError := FALSE;
    wLastStep := WORD#0;
    RETURN;
END_IF

(* ============================================================================
   DECODE ROBOT STATUS (robot -> PLC)
   ============================================================================ *)

(* The job state of the scan we start in (the global transitions below may change it); the
   vw-ks24 decode needs it for the "occupied" term. *)
_bInJob := (_eState = E_RobotState.RS_JOB_WAIT_READY) OR (_eState = E_RobotState.RS_JOB_SEND)
           OR (_eState = E_RobotState.RS_JOB_START) OR (_eState = E_RobotState.RS_JOB_WAIT_RUNNING)
           OR (_eState = E_RobotState.RS_JOB_RUNNING);

IF GVL_Cell.PROFILE_VW THEN
    (* ---- VW KS24 signal map (status bits addressed by $OUT index) ---- *)
    _nIdx := GVL_Cell.VW_READY_OUT;
    _nB := (_nIdx - 1) / 8;
    _nBit := (_nIdx - 1) MOD 8;
    bRobotReady := (SHR(BYTE_TO_WORD(stIn.aVassIn[_nB]), _nBit) AND WORD#1) = WORD#1;

    _nIdx := GVL_Cell.VW_AUTO_OUT;
    _nB := (_nIdx - 1) / 8;
    _nBit := (_nIdx - 1) MOD 8;
    bModeExt := (SHR(BYTE_TO_WORD(stIn.aVassIn[_nB]), _nBit) AND WORD#1) = WORD#1;

    _nIdx := GVL_Cell.VW_PF0_OUT;
    _nB := (_nIdx - 1) / 8;
    _nBit := (_nIdx - 1) MOD 8;
    bAtHome := (SHR(BYTE_TO_WORD(stIn.aVassIn[_nB]), _nBit) AND WORD#1) = WORD#1;

    _nIdx := GVL_Cell.VW_END_OUT;
    _nB := (_nIdx - 1) / 8;
    _nBit := (_nIdx - 1) MOD 8;
    _bFolgeEnd := (SHR(BYTE_TO_WORD(stIn.aVassIn[_nB]), _nBit) AND WORD#1) = WORD#1;
    bProgFinished := _bFolgeEnd;

    (* A10 (RK100: user_saf and em_stop group) is the drive / safety-circuit feedback; A9
       (Bereit) drops while a Folge runs, so it is only used for the job handshake. *)
    _nIdx := GVL_Cell.VW_RK100_OUT;
    _nB := (_nIdx - 1) / 8;
    _nBit := (_nIdx - 1) MOD 8;
    _bTmp := (SHR(BYTE_TO_WORD(stIn.aVassIn[_nB]), _nBit) AND WORD#1) = WORD#1;
    bDrivesOn := _bTmp;
    _nIdx := GVL_Cell.VW_ESTOP_OUT;
    _nB := (_nIdx - 1) / 8;
    _nBit := (_nIdx - 1) MOD 8;
    bSafetyOK := _bTmp AND ((SHR(BYTE_TO_WORD(stIn.aVassIn[_nB]), _nBit) AND WORD#1) = WORD#1)
                 AND stIn.abySafeIn[0].0 AND stIn.abySafeIn[1].4;

    (* Echo: PRG_NR_REFL A1-8 *)
    wActiveJob := BYTE_TO_WORD(stIn.aVassIn[0]);
    bJobAck := (wActiveJob <> WORD#0) AND (wActiveJob = _wJob);

    (* Op index: P_PktNr_SPS, 16 bits little-endian from VW_STEP_OUT *)
    _nB := (GVL_Cell.VW_STEP_OUT - 1) / 8;
    wStep := BYTE_TO_WORD(stIn.aVassIn[_nB]) OR SHL(BYTE_TO_WORD(stIn.aVassIn[_nB + 1]), 8);

    (* Error code: VW_FEH_BIN_A, 8 bits *)
    _nB := (GVL_Cell.VW_ERR_OUT - 1) / 8;
    wRobotErrorCode := BYTE_TO_WORD(stIn.aVassIn[_nB]);
    bRobotError := wRobotErrorCode <> WORD#0;

    (* REQUEST bit z = A(80+n) OR NOT A(40+n): requesting, or inside ("occupied"). The
       release is A(40+n) going TRUE again, which drops the bit. The "occupied" term counts
       only while this driver has a job: an all-zero frame (robot not connected yet, PROFINET
       down) would otherwise read as "inside every interlock". *)
    dwZoneReq := DWORD#0;
    FOR _z := 1 TO GVL_Cell.N_ZONES DO
        _n := GVL_Cell.anInterlock[(nRobot - 1) * GVL_Cell.N_ZONES + _z];
        IF (_n >= 1) AND (_n <= 16) THEN
            _nIdx := GVL_Cell.VW_REQ_OUT + _n - 1;
            _nB := (_nIdx - 1) / 8;
            _nBit := (_nIdx - 1) MOD 8;
            _bTmp := (SHR(BYTE_TO_WORD(stIn.aVassIn[_nB]), _nBit) AND WORD#1) = WORD#1;
            _nIdx := GVL_Cell.VW_REL_OUT + _n - 1;
            _nB := (_nIdx - 1) / 8;
            _nBit := (_nIdx - 1) MOD 8;
            IF _bTmp OR (_bInJob AND ((SHR(BYTE_TO_WORD(stIn.aVassIn[_nB]), _nBit) AND WORD#1) = WORD#0)) THEN
                dwZoneReq := dwZoneReq OR SHL(DWORD#1, _z - 1);
            END_IF
        END_IF
    END_FOR

    (* No ProgRunning bit: the Folge runs while its number is echoed and the robot is neither
       at its home point nor reporting the Folge end. *)
    bProgRunning := (wActiveJob <> WORD#0) AND (wActiveJob = _wJob) AND NOT bAtHome
                    AND NOT _bFolgeEnd;
ELSE
    (* Status word byte 0 / 1 *)
    bDrivesOn     := stIn.aVassIn[0].0;
    bProgRunning  := stIn.aVassIn[0].1;
    bAtHome       := stIn.aVassIn[0].2;
    bModeExt      := stIn.aVassIn[0].4;
    bRobotReady   := stIn.aVassIn[0].5;
    bRobotError   := stIn.aVassIn[0].6;
    bProgFinished := stIn.aVassIn[1].2;
    bJobAck       := stIn.aVassIn[1].3;

    (* Echoed job number from bytes 2-3 (or byte 2 only) *)
    IF GVL_Cell.JOB_NUMBER_BYTE THEN
        wActiveJob := BYTE_TO_WORD(stIn.aVassIn[2]);
    ELSE
        wActiveJob := BYTE_TO_WORD(stIn.aVassIn[2])
                      OR SHL(BYTE_TO_WORD(stIn.aVassIn[3]), 8);
    END_IF

    (* Op index (WORD LE) and zone REQUEST (DWORD LE) *)
    wStep := BYTE_TO_WORD(stIn.aVassIn[GVL_Cell.STEP_BYTE])
             OR SHL(BYTE_TO_WORD(stIn.aVassIn[GVL_Cell.STEP_BYTE + 1]), 8);

    dwZoneReq := BYTE_TO_DWORD(stIn.aVassIn[GVL_Cell.REQ_BYTE])
                 OR SHL(BYTE_TO_DWORD(stIn.aVassIn[GVL_Cell.REQ_BYTE + 1]), 8)
                 OR SHL(BYTE_TO_DWORD(stIn.aVassIn[GVL_Cell.REQ_BYTE + 2]), 16)
                 OR SHL(BYTE_TO_DWORD(stIn.aVassIn[GVL_Cell.REQ_BYTE + 3]), 24);

    (* Error code from bytes 10-11 *)
    wRobotErrorCode := BYTE_TO_WORD(stIn.aVassIn[10])
                       OR SHL(BYTE_TO_WORD(stIn.aVassIn[11]), 8);

    (* Safety status: SafeIn0.0 drives OK, SafeIn1.4 E-Stop OK *)
    bSafetyOK := stIn.abySafeIn[0].0 AND stIn.abySafeIn[1].4;
END_IF

(* SIMULATION ONLY (bt2plc [[robot]] safety_bypass -> GVL_Cell.abSafetyBypass, e.g. a KUKA virtual controller whose FDIO64
   slot carries no F-data to this non-safety controller): the slot-1 bits are not required. The
   vw-ks24 drive / E-stop status bits still count. *)
IF (nRobot >= 1) AND (nRobot <= GVL_Cell.N_ROBOTS) AND GVL_Cell.abSafetyBypass[nRobot] THEN
    IF GVL_Cell.PROFILE_VW THEN
        _nIdx := GVL_Cell.VW_ESTOP_OUT;
        _nB := (_nIdx - 1) / 8;
        _nBit := (_nIdx - 1) MOD 8;
        bSafetyOK := bDrivesOn AND ((SHR(BYTE_TO_WORD(stIn.aVassIn[_nB]), _nBit) AND WORD#1) = WORD#1);
    ELSE
        bSafetyOK := TRUE;
    END_IF
END_IF

(* ============================================================================
   EDGES
   ============================================================================ *)
_rtrigJob(CLK := bCmdJob);
_rtrigReset(CLK := bCmdReset);
IF _rtrigJob.Q THEN
    _bJobPending := TRUE;
END_IF
IF NOT bCmdJob THEN
    _bJobPending := FALSE;
END_IF

(* ============================================================================
   GLOBAL TRANSITIONS
   ============================================================================ *)
_bInJob := (_eState = E_RobotState.RS_JOB_WAIT_READY) OR (_eState = E_RobotState.RS_JOB_SEND)
           OR (_eState = E_RobotState.RS_JOB_START) OR (_eState = E_RobotState.RS_JOB_WAIT_RUNNING)
           OR (_eState = E_RobotState.RS_JOB_RUNNING);
_bUp := _bInJob OR (_eState = E_RobotState.RS_IDLE);
_bNoJob := (_eState = E_RobotState.RS_OFF) OR (_eState = E_RobotState.RS_SAFETY_ENABLE)
           OR (_eState = E_RobotState.RS_DRIVES_ON) OR (_eState = E_RobotState.RS_MODE_EXT)
           OR (_eState = E_RobotState.RS_IDLE);

IF _bInJob AND bCmdStop THEN
    _eState := E_RobotState.RS_STOPPING;
ELSIF _bUp AND bRobotError THEN
    eError := E_CellError.ERR_ROBOT_ERROR;
    _eState := E_RobotState.RS_ERROR;
ELSIF _bUp AND NOT bSafetyOK THEN
    eError := E_CellError.ERR_SAFETY_LOST;
    _eState := E_RobotState.RS_ERROR;
ELSIF _bUp AND NOT bDrivesOn THEN
    eError := E_CellError.ERR_DRIVES_LOST;
    _eState := E_RobotState.RS_ERROR;
ELSIF _bNoJob AND bProgRunning AND NOT GVL_Cell.PROFILE_VW THEN
    (* a program runs that this driver did not start (head restart / download, manual
       start): RS_ERROR holds Stop + Cancel while ProgRunning *)
    eError := E_CellError.ERR_UNEXPECTED_RUN;
    _eState := E_RobotState.RS_ERROR;
END_IF

(* ============================================================================
   STATE TIMER (after the global transitions: a new state always starts with
   fresh timers, also when it was entered by a global transition this scan)
   ============================================================================ *)
IF _eState <> _eLastState THEN
    _tonStep(IN := FALSE);
    _tonPulse(IN := FALSE);
    _tonStopDebounce(IN := FALSE);
    _eLastState := _eState;
END_IF
IF _eState = E_RobotState.RS_STOPPING THEN
    _tStepLimit := GVL_Cell.T_ABORT_LIMIT;
ELSIF _eState = E_RobotState.RS_SAFETY_ENABLE THEN
    _tStepLimit := GVL_Cell.T_BRINGUP_LIMIT;    (* PROFINET / PROFIsafe connection set-up *)
ELSE
    _tStepLimit := GVL_Cell.T_HANDSHAKE;        (* drives / EXT and job handshakes *)
END_IF
_tonStep(IN := TRUE, PT := _tStepLimit);

(* ============================================================================
   STATE MACHINE
   ============================================================================ *)
CASE _eState OF

E_RobotState.RS_OFF:
    _bSafeEnable := FALSE;
    _bDrivesOnCmd := FALSE;
    _bExtCmd := FALSE;
    _bJobReqCmd := FALSE;
    _bStartCmd := FALSE;
    _bStopCmd := FALSE;
    _bCancelCmd := FALSE;
    _bResetCmd := FALSE;
    IF bPowerOn THEN
        _eState := E_RobotState.RS_SAFETY_ENABLE;
    END_IF

E_RobotState.RS_SAFETY_ENABLE:
    _bSafeEnable := TRUE;
    IF bSafetyOK THEN
        _eState := E_RobotState.RS_DRIVES_ON;
    ELSIF _tonStep.Q THEN
        eError := E_CellError.ERR_SAFETY_TIMEOUT;
        _eState := E_RobotState.RS_ERROR;
    END_IF

E_RobotState.RS_DRIVES_ON:
    _bDrivesOnCmd := TRUE;
    IF bDrivesOn THEN
        _eState := E_RobotState.RS_MODE_EXT;
    ELSIF _tonStep.Q THEN
        eError := E_CellError.ERR_DRIVES_TIMEOUT;
        _eState := E_RobotState.RS_ERROR;
    END_IF

E_RobotState.RS_MODE_EXT:
    _bExtCmd := TRUE;
    IF bModeExt THEN
        _eState := E_RobotState.RS_IDLE;
    ELSIF _tonStep.Q THEN
        eError := E_CellError.ERR_EXT_TIMEOUT;
        _eState := E_RobotState.RS_ERROR;
    END_IF

E_RobotState.RS_IDLE:
    _bJobReqCmd := FALSE;
    _bStartCmd := FALSE;
    _bStopCmd := FALSE;
    _bCancelCmd := FALSE;
    IF NOT bCmdJob THEN
        bJobDone := FALSE;
    END_IF
    IF NOT bPowerOn THEN
        _eState := E_RobotState.RS_OFF;
    ELSIF _bJobPending THEN
        _bJobPending := FALSE;
        _wJob := wJobNr;
        _bProdJob := bProdJob;
        bJobDone := FALSE;
        wLastStep := WORD#0;
        _eState := E_RobotState.RS_JOB_WAIT_READY;
    END_IF

E_RobotState.RS_JOB_WAIT_READY:
    _bJobReqCmd := FALSE;                   (* guarantees a rising edge in RS_JOB_SEND *)
    _bVwStarted := FALSE;
    IF GVL_Cell.PROFILE_VW THEN
        (* the robot waits at its home point with PRG_NR_REFL = 0 *)
        IF bRobotReady AND bAtHome AND (wActiveJob = WORD#0) THEN
            _eState := E_RobotState.RS_JOB_SEND;
        ELSIF _tonStep.Q THEN
            eError := E_CellError.ERR_NOT_READY;
            _eState := E_RobotState.RS_ERROR;
        END_IF
    ELSIF bRobotReady AND NOT bJobAck THEN
        _eState := E_RobotState.RS_JOB_SEND;
    ELSIF _tonStep.Q THEN
        eError := E_CellError.ERR_NOT_READY;
        _eState := E_RobotState.RS_ERROR;
    END_IF

E_RobotState.RS_JOB_SEND:
    _bJobReqCmd := TRUE;                    (* vw: PRG_NR is written in the encode section *)
    IF GVL_Cell.PROFILE_VW THEN
        (* the robot mirrors PRG_NR on A1-8 while it waits for the Folge start *)
        IF wActiveJob = _wJob THEN
            _eState := E_RobotState.RS_JOB_START;
        ELSIF _tonStep.Q THEN
            eError := E_CellError.ERR_ACK_TIMEOUT;
            _eState := E_RobotState.RS_ERROR;
        END_IF
    ELSIF bJobAck THEN
        _bJobReqCmd := FALSE;
        IF wActiveJob = _wJob THEN
            _eState := E_RobotState.RS_JOB_START;
        ELSE
            eError := E_CellError.ERR_ECHO_MISMATCH;
            _eState := E_RobotState.RS_ERROR;
        END_IF
    ELSIF _tonStep.Q THEN
        _bJobReqCmd := FALSE;
        eError := E_CellError.ERR_ACK_TIMEOUT;
        _eState := E_RobotState.RS_ERROR;
    END_IF

E_RobotState.RS_JOB_START:
    _bStartCmd := TRUE;
    IF GVL_Cell.PROFILE_VW THEN
        (* SRB stays a level until the robot leaves its home point (its cycle start clears PF0) *)
        _bJobReqCmd := TRUE;                (* keep PRG_NR *)
        IF NOT bAtHome THEN
            _bVwStarted := TRUE;
            _bStartCmd := FALSE;
            _eState := E_RobotState.RS_JOB_RUNNING;
        ELSIF _tonStep.Q THEN
            eError := E_CellError.ERR_START_TIMEOUT;
            _eState := E_RobotState.RS_ERROR;
        END_IF
    ELSE
        _bJobReqCmd := FALSE;
        _tonPulse(IN := TRUE, PT := GVL_Cell.T_START_PULSE);
        IF _tonPulse.Q THEN
            _bStartCmd := FALSE;
            _eState := E_RobotState.RS_JOB_WAIT_RUNNING;
        END_IF
    END_IF

E_RobotState.RS_JOB_WAIT_RUNNING:
    _bStartCmd := FALSE;
    IF bProgRunning THEN
        _eState := E_RobotState.RS_JOB_RUNNING;
    ELSIF bProgFinished THEN
        (* finished between two scans - the robot clears ProgFinished on job accept *)
        _eState := E_RobotState.RS_JOB_DONE;
    ELSIF _tonStep.Q THEN
        eError := E_CellError.ERR_START_TIMEOUT;
        _eState := E_RobotState.RS_ERROR;
    END_IF

E_RobotState.RS_JOB_RUNNING:
    (* no timeout here: per-op watchdogs in FB_Cell, HOME uses T_HOME_LIMIT *)
    IF GVL_Cell.PROFILE_VW THEN
        _bJobReqCmd := TRUE;                (* keep PRG_NR until the Folge end *)
        IF _bFolgeEnd THEN
            _eState := E_RobotState.RS_JOB_DONE;
        END_IF
    ELSE
        (* ProgRunning low without ProgFinished is a stop only when it lasts T_STOP_DEBOUNCE:
           the robot writes the two bits to its outputs one after the other (KRL submit), so a
           bus frame taken between them shows both low for one cycle at a normal Folge end. *)
        _tonStopDebounce(IN := NOT bProgRunning AND NOT bProgFinished, PT := GVL_Cell.T_STOP_DEBOUNCE);
        IF bProgFinished AND NOT bProgRunning THEN
            _eState := E_RobotState.RS_JOB_DONE;
        ELSIF _tonStopDebounce.Q THEN
            eError := E_CellError.ERR_ROBOT_STOPPED;
            _eState := E_RobotState.RS_ERROR;
        END_IF
    END_IF

E_RobotState.RS_JOB_DONE:
    IF GVL_Cell.PROFILE_VW THEN
        (* clear PRG_NR, then wait for the Folge end (A14) to fall before the next job *)
        _bJobReqCmd := FALSE;
        IF NOT _bFolgeEnd THEN
            bJobDone := TRUE;
            _eState := E_RobotState.RS_IDLE;
        ELSIF _tonStep.Q THEN
            eError := E_CellError.ERR_HANDSHAKE;
            _eState := E_RobotState.RS_ERROR;
        END_IF
    ELSE
        bJobDone := TRUE;
        _eState := E_RobotState.RS_IDLE;
    END_IF

E_RobotState.RS_STOPPING:
    _bJobReqCmd := FALSE;                   (* vw: clears PRG_NR; FB_Cell withdraws the grants
                                               and partner releases, which stops the robot on
                                               its path through its own driving condition *)
    _bStartCmd := FALSE;
    _bStopCmd := TRUE;
    _bCancelCmd := TRUE;
    IF GVL_Cell.PROFILE_VW THEN
        _bDrivesOnCmd := FALSE;             (* no Stop/Cancel bits in KS24: drop the drives *)
    END_IF
    _tonPulse(IN := TRUE, PT := GVL_Cell.T_STOP_PULSE);
    IF _tonPulse.Q AND NOT bProgRunning THEN
        _bStopCmd := FALSE;
        _bCancelCmd := FALSE;
        _eState := E_RobotState.RS_IDLE;
    ELSIF _tonStep.Q THEN
        (* keep Stop + Cancel: RS_ERROR holds them while ProgRunning *)
        eError := E_CellError.ERR_STOP_TIMEOUT;
        _eState := E_RobotState.RS_ERROR;
    END_IF

E_RobotState.RS_ERROR:
    _bJobReqCmd := FALSE;
    _bStartCmd := FALSE;
    _bStopCmd := bProgRunning;              (* never drop Stop while the robot still runs *)
    _bCancelCmd := bProgRunning;
    _bResetCmd := FALSE;
    IF _rtrigReset.Q THEN
        _eState := E_RobotState.RS_RESET;
    END_IF

E_RobotState.RS_RESET:
    _bStopCmd := bProgRunning;
    _bCancelCmd := bProgRunning;
    (* DrivesOn low while Reset is held: a KUKA controller switches the drives on only at a rising edge of
       $DRIVES_ON after the messages are acknowledged ($CONF_MESS), so RS_DRIVES_ON must raise it again *)
    _bDrivesOnCmd := FALSE;
    _bResetCmd := TRUE;                     (* held >= 500 ms - robot requirement *)
    _tonPulse(IN := TRUE, PT := GVL_Cell.T_RESET_PULSE);
    IF NOT bCmdReset THEN
        (* reset withdrawn by the cell (operator stop): Reset low, error kept *)
        _bResetCmd := FALSE;
        _eState := E_RobotState.RS_ERROR;
    ELSIF _tonPulse.Q THEN
        _bResetCmd := FALSE;
        IF bProgRunning THEN
            (* never leave the error with a running program: RS_ERROR keeps Stop + Cancel *)
            eError := E_CellError.ERR_STOP_TIMEOUT;
            _eState := E_RobotState.RS_ERROR;
        ELSIF NOT bRobotError THEN
            eError := E_CellError.ERR_NONE;
            _eState := E_RobotState.RS_SAFETY_ENABLE;
        ELSE
            eError := E_CellError.ERR_RESET_FAILED;
            _eState := E_RobotState.RS_ERROR;
        END_IF
    END_IF

END_CASE

(* ============================================================================
   JOB STATUS
   ============================================================================ *)
_bInJob := (_eState = E_RobotState.RS_JOB_WAIT_READY) OR (_eState = E_RobotState.RS_JOB_SEND)
           OR (_eState = E_RobotState.RS_JOB_START) OR (_eState = E_RobotState.RS_JOB_WAIT_RUNNING)
           OR (_eState = E_RobotState.RS_JOB_RUNNING);
bJobActive := bProgRunning AND ((_eState = E_RobotState.RS_JOB_START)
              OR (_eState = E_RobotState.RS_JOB_WAIT_RUNNING) OR (_eState = E_RobotState.RS_JOB_RUNNING));

(* Latched max op index of the running production job (step 0 = between jobs) *)
IF bJobActive AND _bProdJob AND (wStep > wLastStep) THEN
    wLastStep := wStep;
END_IF

(* ============================================================================
   ENCODE COMMANDS (PLC -> robot)
   ============================================================================ *)
IF GVL_Cell.PROFILE_VW THEN
    (* ---- VW KS24 commands: PRG_NR A1-8, SRB, drives, acknowledge ---- *)
    FOR _i := 0 TO 31 DO
        stOut.aVassOut[_i] := BYTE#0;
    END_FOR
    (* PRG_NR only from RS_JOB_SEND on: in RS_JOB_WAIT_READY the robot must still echo 0
       (it picks the number up through cell.src as soon as it is written). *)
    IF _bJobReqCmd THEN
        stOut.aVassOut[0] := WORD_TO_BYTE(_wJob AND WORD#16#FF);
    END_IF
    _nIdx := GVL_Cell.VW_SRB_IN;
    _nB := (_nIdx - 1) / 8;
    _nBit := (_nIdx - 1) MOD 8;
    IF _bStartCmd THEN
        _wTmp := BYTE_TO_WORD(stOut.aVassOut[_nB]) OR SHL(WORD#1, _nBit);
        stOut.aVassOut[_nB] := WORD_TO_BYTE(_wTmp);
    END_IF
    _nIdx := GVL_Cell.VW_DRIVES_IN;
    _nB := (_nIdx - 1) / 8;
    _nBit := (_nIdx - 1) MOD 8;
    IF _bDrivesOnCmd THEN
        _wTmp := BYTE_TO_WORD(stOut.aVassOut[_nB]) OR SHL(WORD#1, _nBit);
        stOut.aVassOut[_nB] := WORD_TO_BYTE(_wTmp);
    END_IF
    _nIdx := GVL_Cell.VW_RESET_IN;
    _nB := (_nIdx - 1) / 8;
    _nBit := (_nIdx - 1) MOD 8;
    IF _bResetCmd THEN
        _wTmp := BYTE_TO_WORD(stOut.aVassOut[_nB]) OR SHL(WORD#1, _nBit);
        stOut.aVassOut[_nB] := WORD_TO_BYTE(_wTmp);
    END_IF
    (* PLAN_ID on a free telegram byte pair, only with the production job (0 = no check) *)
    IF (GVL_Cell.PLAN_ID_BYTE > 0) AND _bInJob AND _bProdJob THEN
        stOut.aVassOut[GVL_Cell.PLAN_ID_BYTE]     := WORD_TO_BYTE(GVL_Cell.PLAN_ID AND WORD#16#FF);
        stOut.aVassOut[GVL_Cell.PLAN_ID_BYTE + 1] := WORD_TO_BYTE(SHR(GVL_Cell.PLAN_ID, 8) AND WORD#16#FF);
    END_IF
    (* The interlock grants E(80+n) and partner releases E(40+n) are written by FB_Cell. *)
ELSE
stOut.aVassOut[0].0 := _bDrivesOnCmd;
stOut.aVassOut[0].1 := _bStartCmd;
stOut.aVassOut[0].2 := _bStopCmd;
stOut.aVassOut[0].3 := _bCancelCmd;
stOut.aVassOut[0].4 := _bExtCmd;
stOut.aVassOut[0].5 := _bResetCmd;
stOut.aVassOut[0].6 := FALSE;               (* homing uses HOME_FOLGE, not HomeRequest *)
(* MoveEnable: held in every state but RS_OFF, also through a reset (DrivesOn drops there for the
   $DRIVES_ON edge). A KUKA KSS 9.2 maps $MOVE_ENABLE to it: it refuses EXT with $MOVE_ENABLE on the
   always-TRUE $IN[1025] (M_249), and a motion enable that dropped with DrivesOn needs a new
   acknowledgement (M_1210) before the drives come on. The robot simulator ignores this bit. *)
stOut.aVassOut[0].7 := _eState <> E_RobotState.RS_OFF;
stOut.aVassOut[1].0 := _bJobReqCmd;

(* Job number, bytes 2-3 (or byte 2 only) *)
IF _bInJob THEN
    stOut.aVassOut[2] := WORD_TO_BYTE(_wJob AND WORD#16#FF);
    IF GVL_Cell.JOB_NUMBER_BYTE THEN
        stOut.aVassOut[3] := BYTE#0;
    ELSE
        stOut.aVassOut[3] := WORD_TO_BYTE(SHR(_wJob, 8) AND WORD#16#FF);
    END_IF
ELSE
    stOut.aVassOut[2] := BYTE#0;
    stOut.aVassOut[3] := BYTE#0;
END_IF

(* PLAN_ID, only with the production job *)
IF _bInJob AND _bProdJob THEN
    stOut.aVassOut[GVL_Cell.PLAN_ID_BYTE]     := WORD_TO_BYTE(GVL_Cell.PLAN_ID AND WORD#16#FF);
    stOut.aVassOut[GVL_Cell.PLAN_ID_BYTE + 1] := WORD_TO_BYTE(SHR(GVL_Cell.PLAN_ID, 8) AND WORD#16#FF);
ELSE
    stOut.aVassOut[GVL_Cell.PLAN_ID_BYTE]     := BYTE#0;
    stOut.aVassOut[GVL_Cell.PLAN_ID_BYTE + 1] := BYTE#0;
END_IF

(* GRANT bytes: encoded by FB_Cell after FB_ZoneArbiter *)
stOut.aVassOut[GVL_Cell.GRANT_BYTE]     := BYTE#0;
stOut.aVassOut[GVL_Cell.GRANT_BYTE + 1] := BYTE#0;
stOut.aVassOut[GVL_Cell.GRANT_BYTE + 2] := BYTE#0;
stOut.aVassOut[GVL_Cell.GRANT_BYTE + 3] := BYTE#0;
END_IF

(* Safe outputs *)
IF _bSafeEnable THEN
    stOut.abySafeOut[0] := BYTE#16#01;      (* drive enable *)
    stOut.abySafeOut[1] := BYTE#16#0F;      (* zones 1-4 enable *)
ELSE
    stOut.abySafeOut[0] := BYTE#0;
    stOut.abySafeOut[1] := BYTE#0;
END_IF

(* ============================================================================
   PUBLISH
   ============================================================================ *)
eState := _eState;
bIdle  := (_eState = E_RobotState.RS_IDLE);
bBusy  := _bInJob OR (_eState = E_RobotState.RS_STOPPING) OR (_eState = E_RobotState.RS_RESET);
bError := (_eState = E_RobotState.RS_ERROR) OR (_eState = E_RobotState.RS_RESET);

(* ---- FB_ZoneArbiter_Body.st ---- *)
(*
 * FB_ZoneArbiter - Implementation
 * Order per scan: debounce + handshake check, release, grant, fault latch.
 *)

IF bReset THEN
    FOR _z := 1 TO GVL_Cell.N_ZONES DO
        anHolder[_z] := 0;
        anTicket[_z] := GVL_Cell.anZoneFirst[_z];
    END_FOR
    FOR _r := 1 TO GVL_Cell.N_ROBOTS DO
        adwGrant[_r] := DWORD#0;
        _audiWaitSince[_r] := 0;
        _anGrantStep[_r] := 0;
        _awPrevStep[_r] := awStep[_r];
        _adwPrevReq[_r] := adwReq[_r];
        _atChange[_r] := tNow;
        _abStable[_r] := FALSE;
    END_FOR
    _udiScan := 0;
    bFault := FALSE;
    eFault := E_CellError.ERR_NONE;
    nFaultRobot := 0;
    nFaultZone := 0;
    bAllConsumed := (GVL_Cell.N_ZONES = 0) OR (ePolicy = E_GrantPolicy.GP_FCFS);
    RETURN;
END_IF

IF bFault THEN
    RETURN;                                 (* latched until bReset *)
END_IF

_udiScan := _udiScan + 1;
_eNew := E_CellError.ERR_NONE;
_nNewRobot := 0;
_nNewZone := 0;

(* ============================================================================
   0. DEBOUNCE / 4-PHASE HANDSHAKE
   ============================================================================ *)
FOR _r := 1 TO GVL_Cell.N_ROBOTS DO
    IF (awStep[_r] <> _awPrevStep[_r]) OR (adwReq[_r] <> _adwPrevReq[_r]) THEN
        _atChange[_r] := tNow;
        _awPrevStep[_r] := awStep[_r];
        _adwPrevReq[_r] := adwReq[_r];
    END_IF
    _abStable[_r] := (tNow - _atChange[_r]) >= tDebounce;

    (* A correct robot changes its op index only after it has seen GRANT = 0. Profile vw-ks24
       has no 4-phase handshake: there the robot only holds its release level long enough for
       the head to see it (bt2krl emits a dwell after every release), so the check needs the
       debounce to avoid firing on scan jitter. *)
    IF (adwGrant[_r] <> DWORD#0) AND (WORD_TO_INT(awStep[_r]) <> _anGrantStep[_r])
       AND (_abStable[_r] OR NOT GVL_Cell.PROFILE_VW)
       AND (_eNew = E_CellError.ERR_NONE) THEN
        _eNew := E_CellError.ERR_HANDSHAKE;
        _nNewRobot := _r;
        _nNewZone := 0;
    END_IF
END_FOR

(* ============================================================================
   1. RELEASE - holder dropped its REQUEST bit
   ============================================================================ *)
FOR _z := 1 TO GVL_Cell.N_ZONES DO
    _rr := anHolder[_z];
    IF _rr <> 0 THEN
        _dwBit := SHL(DWORD#1, _z - 1);
        IF (adwReq[_rr] AND _dwBit) = DWORD#0 THEN
            IF abRobotOk[_rr] THEN
                anHolder[_z] := 0;
                adwGrant[_rr] := adwGrant[_rr] AND NOT _dwBit;
                IF ePolicy = E_GrantPolicy.GP_PLANNED THEN
                    anTicket[_z] := anTicket[_z] + 1;
                END_IF
            ELSIF _eNew = E_CellError.ERR_NONE THEN
                (* request vanished because the robot stopped / faulted / lost
                   connection: the zone may still be occupied - never re-grant *)
                _eNew := E_CellError.ERR_RELEASE_INVALID;
                _nNewRobot := _rr;
                _nNewZone := _z;
            END_IF
        END_IF
    END_IF
END_FOR

(* Permit bit: not a mutex, released as soon as REQUEST bit 31 drops *)
FOR _r := 1 TO GVL_Cell.N_ROBOTS DO
    IF ((adwGrant[_r] AND GVL_Cell.PERMIT_MASK) <> DWORD#0)
       AND ((adwReq[_r] AND GVL_Cell.PERMIT_MASK) = DWORD#0) THEN
        adwGrant[_r] := adwGrant[_r] AND NOT GVL_Cell.PERMIT_MASK;
    END_IF
END_FOR

(* ============================================================================
   2. GRANT
   ============================================================================ *)
FOR _r := 1 TO GVL_Cell.N_ROBOTS DO
    _abPicked[_r] := FALSE;
    IF (adwReq[_r] = DWORD#0) OR (adwGrant[_r] <> DWORD#0) THEN
        _audiWaitSince[_r] := 0;
    ELSIF _audiWaitSince[_r] = 0 THEN
        _audiWaitSince[_r] := _udiScan;
    END_IF
END_FOR
_dwReserved := DWORD#0;

FOR _k := 1 TO GVL_Cell.N_ROBOTS DO
    (* --- visiting order: PLANNED = robot index, FCFS = oldest request first --- *)
    _rSel := 0;
    FOR _r := 1 TO GVL_Cell.N_ROBOTS DO
        IF NOT _abPicked[_r] THEN
            IF _rSel = 0 THEN
                _rSel := _r;
            ELSIF (ePolicy = E_GrantPolicy.GP_FCFS) AND (_audiWaitSince[_r] <> 0) THEN
                IF (_audiWaitSince[_rSel] = 0) OR (_audiWaitSince[_r] < _audiWaitSince[_rSel]) THEN
                    _rSel := _r;
                END_IF
            END_IF
        END_IF
    END_FOR
    _rr := _rSel;
    _abPicked[_rr] := TRUE;

    (* --- expected mask of the op the robot reports --- *)
    _nStep := WORD_TO_INT(awStep[_rr]);
    _iOp := 0;
    _dwExp := DWORD#0;
    IF (_nStep >= 1) AND (_nStep <= GVL_Cell.anRobotOpCount[_rr]) THEN
        _iOp := GVL_Cell.anRobotFirstOp[_rr] + _nStep - 1;
        _dwExp := GVL_Cell.aOps[_iOp].dwZoneMask;
    END_IF
    _dwZones := _dwExp AND NOT GVL_Cell.PERMIT_MASK;

    _bPending := bEnable AND abRobotOk[_rr] AND (adwReq[_rr] <> DWORD#0) AND (adwGrant[_rr] = DWORD#0);

    (* --- request must equal the op mask (debounced) --- *)
    IF _bPending AND _abStable[_rr] AND (adwReq[_rr] <> _dwExp)
       AND (_eNew = E_CellError.ERR_NONE) THEN
        _eNew := E_CellError.ERR_REQ_MISMATCH;
        _nNewRobot := _rr;
        _nNewZone := 0;
    END_IF

    (* --- a holder must not raise bits it was not granted --- *)
    IF (adwGrant[_rr] <> DWORD#0) AND ((adwReq[_rr] AND NOT adwGrant[_rr]) <> DWORD#0)
       AND (_eNew = E_CellError.ERR_NONE) THEN
        _eNew := E_CellError.ERR_UNEXPECTED_REQUEST;
        _nNewRobot := _rr;
        _nNewZone := 0;
    END_IF

    IF _bPending AND (adwReq[_rr] = _dwExp) THEN
        (* --- zones: all free, (planned) ticket = this op, (FCFS) not reserved --- *)
        _bOk := TRUE;
        FOR _z := 1 TO GVL_Cell.N_ZONES DO
            _dwBit := SHL(DWORD#1, _z - 1);
            IF (_dwZones AND _dwBit) <> DWORD#0 THEN
                IF anHolder[_z] <> 0 THEN
                    _bOk := FALSE;
                ELSIF ePolicy = E_GrantPolicy.GP_PLANNED THEN
                    _nTicket := anTicket[_z];
                    _nLastTicket := GVL_Cell.anZoneFirst[_z] + GVL_Cell.anZoneCount[_z] - 1;
                    IF (_nTicket < GVL_Cell.anZoneFirst[_z]) OR (_nTicket > _nLastTicket) THEN
                        _bOk := FALSE;              (* zone consumed *)
                        IF _abStable[_rr] AND (_eNew = E_CellError.ERR_NONE) THEN
                            _eNew := E_CellError.ERR_TICKET_SKIPPED;
                            _nNewRobot := _rr;
                            _nNewZone := _z;
                        END_IF
                    ELSIF (GVL_Cell.aTickets[_nTicket].nRobot <> _rr)
                          OR (GVL_Cell.aTickets[_nTicket].nOp <> _nStep) THEN
                        _bOk := FALSE;              (* not this op's turn yet *)
                        IF (GVL_Cell.aTickets[_nTicket].nRobot = _rr) AND _abStable[_rr]
                           AND (_eNew = E_CellError.ERR_NONE) THEN
                            _eNew := E_CellError.ERR_TICKET_SKIPPED;
                            _nNewRobot := _rr;
                            _nNewZone := _z;
                        END_IF
                    END_IF
                ELSIF (_dwReserved AND _dwBit) <> DWORD#0 THEN
                    _bOk := FALSE;                  (* FCFS: reserved by an older requester *)
                END_IF
            END_IF
        END_FOR

        (* --- permit: every predecessor op done --- *)
        _bPermitOk := TRUE;
        IF ((_dwExp AND GVL_Cell.PERMIT_MASK) <> DWORD#0) AND (_iOp >= 1) THEN
            (* GVL array elements are copied to locals before use as call arguments *)
            _nPredFirst := GVL_Cell.aOps[_iOp].nPredFirst;
            _nPredLast := _nPredFirst + GVL_Cell.aOps[_iOp].nPredCount - 1;
            _nPredFirst := MAX(1, _nPredFirst);
            _nPredLast := MIN(GVL_Cell.N_PREDS, _nPredLast);
            FOR _p := _nPredFirst TO _nPredLast DO
                _q := GVL_Cell.aPreds[_p].nRobot;
                IF (_q < 1) OR (_q > GVL_Cell.N_ROBOTS) THEN
                    _bPermitOk := FALSE;
                ELSIF anDone[_q] < GVL_Cell.aPreds[_p].nOp THEN
                    _bPermitOk := FALSE;
                END_IF
            END_FOR
        END_IF

        IF _bOk AND _bPermitOk THEN
            FOR _z := 1 TO GVL_Cell.N_ZONES DO
                IF (_dwZones AND SHL(DWORD#1, _z - 1)) <> DWORD#0 THEN
                    anHolder[_z] := _rr;
                END_IF
            END_FOR
            adwGrant[_rr] := _dwExp;
            _anGrantStep[_rr] := _nStep;
            _audiWaitSince[_rr] := 0;
        ELSIF _bPermitOk AND (ePolicy = E_GrantPolicy.GP_FCFS) THEN
            (* older requester blocked only by occupied / reserved zones: reserve them
               (a requester still waiting for its permit reserves nothing - no deadlock) *)
            _dwReserved := _dwReserved OR _dwZones;
        END_IF
    END_IF
END_FOR

(* ============================================================================
   3. FAULT LATCH / CYCLE COMPLETENESS
   ============================================================================ *)
IF _eNew <> E_CellError.ERR_NONE THEN
    bFault := TRUE;
    eFault := _eNew;
    nFaultRobot := _nNewRobot;
    nFaultZone := _nNewZone;
    FOR _r := 1 TO GVL_Cell.N_ROBOTS DO
        adwGrant[_r] := DWORD#0;
    END_FOR
END_IF

bAllConsumed := TRUE;
FOR _z := 1 TO GVL_Cell.N_ZONES DO
    IF anHolder[_z] <> 0 THEN
        bAllConsumed := FALSE;
    ELSIF (ePolicy = E_GrantPolicy.GP_PLANNED)
          AND (anTicket[_z] <= GVL_Cell.anZoneFirst[_z] + GVL_Cell.anZoneCount[_z] - 1) THEN
        bAllConsumed := FALSE;
    END_IF
END_FOR

(* ---- PLC_PRG.st ---- *)
(*
 * PLC_PRG - Head PLC cell program
 * Generated by bt2plc 0.1.0 for cell welding_cell_2_small (plan bt_1790934549_welding_cell_2_small)
 *
 * Copies every robot's GVL_IO block into the cell's input array, runs FB_Cell and
 * copies the commands back (whole arrays / single bytes only).
 *
 * Operator (plain VARs, pulses are cleared after each scan):
 *   bAutoRun          Level: start a cycle whenever the cell is READY
 *                     (initialised from GVL_Cell.AUTO_RUN on the first scan)
 *   bStart            Pulse: start one cycle
 *   bStop             Pulse: abort (ERR_OPERATOR_STOP); latched in every state, also
 *                     cancels a running reset (CS_RESETTING -> CS_ERROR)
 *   bReset            Pulse: reset after an error (a pulse during CS_ABORTING is kept)
 *   bRecoveryConfirm  Pulse: after an abort mid-cycle or a start-up with an active robot
 *                     away from home, robots moved clear -> sequential blind homing
 *
 * Status: PLC_PRG.fbCell.eState / eError / nErrorRobot / nErrorOp / nErrorZone /
 *         bRecoveryRequired / udiCycles / tLastCycle / aeRobotState / awStep / adwGrant ...
 *
 * Task: MainTask (4 ms cycle)
 *)

PROGRAM PLC_PRG
VAR
    (* Cell controller *)
    fbCell              : FB_Cell;

    (* === Operator === *)
    bAutoRun            : BOOL := TRUE;     (* overwritten by GVL_Cell.AUTO_RUN on the first scan *)
    bStart              : BOOL;
    bStop               : BOOL;
    bReset              : BOOL;
    bRecoveryConfirm    : BOOL;

    (* === Status readback === *)
    eCellState          : E_CellState;
    eCellError          : E_CellError;
    bCellError          : BOOL;
    bRecoveryRequired   : BOOL;
    udiCycles           : UDINT;

    (* Robot input images for fbCell *)
    _astIn              : ARRAY[1..2] OF ST_RobotIn;
    _bFirstScan         : BOOL := TRUE;
END_VAR

(* ---- PLC_PRG_Body.st ---- *)
(*
 * PLC_PRG - Implementation
 *)

IF _bFirstScan THEN
    bAutoRun := GVL_Cell.AUTO_RUN;
    _bFirstScan := FALSE;
END_IF

(* ============================================================================
   INPUTS: GVL_IO -> fbCell (robot -> PLC)
   ============================================================================ *)

(* 1: R1 - robot1 - kuka_robi1 (kuka-robi1, 192.168.100.11) *)
_astIn[1].abySafeIn[0] := GVL_IO.bySafeIn0_R1;
_astIn[1].abySafeIn[1] := GVL_IO.bySafeIn1_R1;
_astIn[1].abySafeIn[2] := GVL_IO.bySafeIn2_R1;
_astIn[1].abySafeIn[3] := GVL_IO.bySafeIn3_R1;
_astIn[1].abySafeIn[4] := GVL_IO.bySafeIn4_R1;
_astIn[1].abySafeIn[5] := GVL_IO.bySafeIn5_R1;
_astIn[1].abySafeIn[6] := GVL_IO.bySafeIn6_R1;
_astIn[1].abySafeIn[7] := GVL_IO.bySafeIn7_R1;
_astIn[1].aVassIn := GVL_IO.aVassInputData_R1;

(* 2: R2 - robot2 - kuka_robi2 (kuka-robi2, 192.168.100.12) *)
_astIn[2].abySafeIn[0] := GVL_IO.bySafeIn0_R2;
_astIn[2].abySafeIn[1] := GVL_IO.bySafeIn1_R2;
_astIn[2].abySafeIn[2] := GVL_IO.bySafeIn2_R2;
_astIn[2].abySafeIn[3] := GVL_IO.bySafeIn3_R2;
_astIn[2].abySafeIn[4] := GVL_IO.bySafeIn4_R2;
_astIn[2].abySafeIn[5] := GVL_IO.bySafeIn5_R2;
_astIn[2].abySafeIn[6] := GVL_IO.bySafeIn6_R2;
_astIn[2].abySafeIn[7] := GVL_IO.bySafeIn7_R2;
_astIn[2].aVassIn := GVL_IO.aVassInputData_R2;

(* ============================================================================
   CELL
   ============================================================================ *)
fbCell(
    bEnable             := TRUE,
    bAutoRun            := bAutoRun,
    bStart              := bStart,
    bStop               := bStop,
    bReset              := bReset,
    bRecoveryConfirm    := bRecoveryConfirm,
    astIn               := _astIn,
    eState              => eCellState,
    eError              => eCellError,
    bError              => bCellError,
    bRecoveryRequired   => bRecoveryRequired,
    udiCycles           => udiCycles);

(* ============================================================================
   OUTPUTS: fbCell -> GVL_IO (PLC -> robot)
   ============================================================================ *)

(* 1: R1 - robot1 *)
GVL_IO.bySafeOut0_R1 := fbCell.astOut[1].abySafeOut[0];
GVL_IO.bySafeOut1_R1 := fbCell.astOut[1].abySafeOut[1];
GVL_IO.bySafeOut2_R1 := fbCell.astOut[1].abySafeOut[2];
GVL_IO.bySafeOut3_R1 := fbCell.astOut[1].abySafeOut[3];
GVL_IO.bySafeOut4_R1 := fbCell.astOut[1].abySafeOut[4];
GVL_IO.bySafeOut5_R1 := fbCell.astOut[1].abySafeOut[5];
GVL_IO.bySafeOut6_R1 := fbCell.astOut[1].abySafeOut[6];
GVL_IO.bySafeOut7_R1 := fbCell.astOut[1].abySafeOut[7];
GVL_IO.aVassOutputData_R1 := fbCell.astOut[1].aVassOut;

(* 2: R2 - robot2 *)
GVL_IO.bySafeOut0_R2 := fbCell.astOut[2].abySafeOut[0];
GVL_IO.bySafeOut1_R2 := fbCell.astOut[2].abySafeOut[1];
GVL_IO.bySafeOut2_R2 := fbCell.astOut[2].abySafeOut[2];
GVL_IO.bySafeOut3_R2 := fbCell.astOut[2].abySafeOut[3];
GVL_IO.bySafeOut4_R2 := fbCell.astOut[2].abySafeOut[4];
GVL_IO.bySafeOut5_R2 := fbCell.astOut[2].abySafeOut[5];
GVL_IO.bySafeOut6_R2 := fbCell.astOut[2].abySafeOut[6];
GVL_IO.bySafeOut7_R2 := fbCell.astOut[2].abySafeOut[7];
GVL_IO.aVassOutputData_R2 := fbCell.astOut[2].aVassOut;

(* One-shot operator buttons *)
bStart := FALSE;
bStop := FALSE;
bReset := FALSE;
bRecoveryConfirm := FALSE;
